// TwinCAT 3 PLC project TestRunner
// Title: TestRunner
// Company: Intecre Ltd
// ProjectVersion: 1.0.0.0
// Description: TcUnit test suites for the Intecre.Utilities library. Not a library; activate it on a runtime (the usermode runtime works) to run the tests.
// ProgramVersion: 3.1.4026.25
// libraries:
//   Tc2_Standard, * (Beckhoff Automation GmbH)
//   Tc2_System, * (Beckhoff Automation GmbH)
//   Tc2_Utilities, * (Beckhoff Automation GmbH)
//   TcUnit, * (www.tcunit.org)
//   Intecre.Utilities, * (Intecre Ltd)
// project tree:
//   / MAIN.TcPOU, PlcTask.TcTTO, SlowTask.TcTTO, ControllersInSlowTask.TcPOU
//   Tests/ CharIsNumber_Tests.TcPOU, TryStringToDint_Tests.TcPOU, TryStringToUdint_Tests.TcPOU, TryStringToWord_Tests.TcPOU, TryStringToLreal_Tests.TcPOU, F_Concat_Tests.TcPOU, F_ConcatLarge_Tests.TcPOU, F_Gate_Tests.TcPOU, FB_StringList_Tests.TcPOU, FB_UdintList_Tests.TcPOU, FB_PointerList_Tests.TcPOU, FB_LongStringList_Tests.TcPOU, FB_TargList_Tests.TcPOU, FB_Dictionary_Tests.TcPOU, F_DictionaryValuesCrc_Tests.TcPOU, FB_AlphaBetaFilter_Tests.TcPOU, FB_P_Control_Tests.TcPOU, FB_I_Controller_Tests.TcPOU, FB_PI_Controller_Tests.TcPOU, T_Task_Tests.TcPOU, T_NamedBase_Tests.TcPOU, Logger_Tests.TcPOU, FB_Assert_Tests.TcPOU, F_GetKL306xState_Tests.TcPOU, ProjectInformation_Tests.TcPOU, F_TargToString_Tests.TcPOU, F_StringToTarg_Tests.TcPOU, F_GetAmsNetId_Tests.TcPOU, T_Timer_Tests.TcPOU, T_GetHandle_Tests.TcPOU, T_InvokeRpcMethod_Tests.TcPOU, T_WritePersistentData_Tests.TcPOU
//   Mocks/ T_MockExternalLogger.TcPOU, T_RpcTarget.TcPOU, ST_RpcAddParams.TcDUT
// (motion and I/O tree: see PLC project intecreutilities)
// real-time tasks:
//   TASK PlcTask: cycle T#10ms, priority 20, ADS port 350
//   TASK SlowTask: cycle T#50000us, priority 25, ADS port 351

CONFIGURATION TestRunner
    RESOURCE PLC ON TwinCAT3
        TASK PlcTask(INTERVAL := T#10ms, PRIORITY := 20);
        TASK SlowTask(INTERVAL := T#50000us, PRIORITY := 25);
        PROGRAM MAIN WITH PlcTask : MAIN;
        PROGRAM ControllersInSlowTask WITH SlowTask : ControllersInSlowTask;
    END_RESOURCE
END_CONFIGURATION

// ---- Mocks/ST_RpcAddParams.TcDUT
// Input block of T_RpcTarget.Add as sent over ADS.
TYPE ST_RpcAddParams :
STRUCT
  a : DINT;
  b : DINT;
END_STRUCT
END_TYPE

// ---- MAIN.TcPOU
// Runs every TcUnit suite of the Intecre.Utilities library, one suite at a time.
PROGRAM MAIN
VAR
  suiteCharIsNumber        : CharIsNumber_Tests;
  suiteTryStringToDint     : TryStringToDint_Tests;
  suiteTryStringToUdint    : TryStringToUdint_Tests;
  suiteTryStringToWord     : TryStringToWord_Tests;
  suiteTryStringToLreal    : TryStringToLreal_Tests;
  suiteConcat              : F_Concat_Tests;
  suiteConcatLarge         : F_ConcatLarge_Tests;
  suiteGate                : F_Gate_Tests;
  suiteStringList          : FB_StringList_Tests;
  suiteUdintList           : FB_UdintList_Tests;
  suitePointerList         : FB_PointerList_Tests;
  suiteLongStringList      : FB_LongStringList_Tests;
  suiteTargList            : FB_TargList_Tests;
  suiteDictionary          : FB_Dictionary_Tests;
  suiteDictionaryValuesCrc : F_DictionaryValuesCrc_Tests;
  suiteAlphaBetaFilter     : FB_AlphaBetaFilter_Tests;
  suiteP_Control           : FB_P_Control_Tests;
  suiteI_Controller        : FB_I_Controller_Tests;
  suitePI_Controller       : FB_PI_Controller_Tests;
  suiteTask                : T_Task_Tests;
  suiteNamedBase           : T_NamedBase_Tests;
  suiteLogger              : Logger_Tests;
  suiteAssert              : FB_Assert_Tests;
  suiteGetKL306xState      : F_GetKL306xState_Tests;
  suiteProjectInformation  : ProjectInformation_Tests;
  suiteTargToString        : F_TargToString_Tests;
  suiteStringToTarg        : F_StringToTarg_Tests;
  suiteGetAmsNetId         : F_GetAmsNetId_Tests;
  suiteTimer               : T_Timer_Tests;
  suiteGetHandle           : T_GetHandle_Tests;
  suiteInvokeRpc           : T_InvokeRpcMethod_Tests;
  suiteWritePersistentData : T_WritePersistentData_Tests;
END_VAR

TcUnit.RUN_IN_SEQUENCE();

END_PROGRAM

// ---- Tests/CharIsNumber_Tests.TcPOU
FUNCTION_BLOCK CharIsNumber_Tests EXTENDS TcUnit.FB_TestSuite

Test_DigitsAreNumbers();
Test_NonDigitsAreNotNumbers();
Test_MinusAcceptedOnlyByOrMinus();
Test_PeriodAcceptedOnlyByOrPeriod();

METHOD PRIVATE Test_DigitsAreNumbers
VAR
  ch : BYTE;
  allDigits : BOOL := TRUE;
END_VAR
TcUnit.TEST(__POUNAME());

// arrange / act
FOR ch := 48 TO 57 DO
  allDigits := allDigits AND CharIsNumber(ch);
END_FOR

// assert
AssertTrue(Condition := allDigits, Message := 'ASCII 0-9 are numbers');

TEST_FINISHED_NAMED(__POUNAME());
END_METHOD

METHOD PRIVATE Test_NonDigitsAreNotNumbers
TcUnit.TEST(__POUNAME());

// act / assert
AssertFalse(Condition := CharIsNumber(47), Message := 'slash (47) is not a number');
AssertFalse(Condition := CharIsNumber(58), Message := 'colon (58) is not a number');
AssertFalse(Condition := CharIsNumber(65), Message := 'A is not a number');
AssertFalse(Condition := CharIsNumber(32), Message := 'space is not a number');
AssertFalse(Condition := CharIsNumber(45), Message := 'minus is not a number');
AssertFalse(Condition := CharIsNumber(46), Message := 'period is not a number');

TEST_FINISHED_NAMED(__POUNAME());
END_METHOD

METHOD PRIVATE Test_MinusAcceptedOnlyByOrMinus
TcUnit.TEST(__POUNAME());

// act / assert
AssertTrue(Condition := CharIsNumberOrMinus(45), Message := 'minus accepted');
AssertTrue(Condition := CharIsNumberOrMinus(53), Message := 'digit 5 accepted');
AssertFalse(Condition := CharIsNumberOrMinus(46), Message := 'period rejected');
AssertFalse(Condition := CharIsNumberOrMinus(65), Message := 'letter rejected');

TEST_FINISHED_NAMED(__POUNAME());
END_METHOD

METHOD PRIVATE Test_PeriodAcceptedOnlyByOrPeriod
TcUnit.TEST(__POUNAME());

// act / assert
AssertTrue(Condition := CharIsNumberOrPeriod(46), Message := 'period accepted');
AssertTrue(Condition := CharIsNumberOrPeriod(48), Message := 'digit 0 accepted');
AssertFalse(Condition := CharIsNumberOrPeriod(45), Message := 'minus rejected');
AssertFalse(Condition := CharIsNumberOrPeriod(65), Message := 'letter rejected');

TEST_FINISHED_NAMED(__POUNAME());
END_METHOD

END_FUNCTION_BLOCK

// ---- Tests/TryStringToDint_Tests.TcPOU
FUNCTION_BLOCK TryStringToDint_Tests EXTENDS TcUnit.FB_TestSuite

Test_ParsesPositive();
Test_ParsesNegative();
Test_ParsesMaxValue();
Test_RejectsLetters();
Test_RejectsEmptyString();
Test_RejectsMinusInsideNumber();
Test_RejectsPlusSign();

METHOD PRIVATE Test_ParsesPositive
VAR
  value : DINT;
  ok : BOOL;
END_VAR
TcUnit.TEST(__POUNAME());

// act
ok := TryStringToDint('123', value);

// assert
AssertTrue(Condition := ok, Message := '123 parses');
AssertEquals_DINT(Expected := 123, Actual := value, Message := 'parsed value');

TEST_FINISHED_NAMED(__POUNAME());
END_METHOD

METHOD PRIVATE Test_ParsesNegative
VAR
  value : DINT;
  ok : BOOL;
END_VAR
TcUnit.TEST(__POUNAME());

// act
ok := TryStringToDint('-45', value);

// assert
AssertTrue(Condition := ok, Message := '-45 parses');
AssertEquals_DINT(Expected := -45, Actual := value, Message := 'parsed value');

TEST_FINISHED_NAMED(__POUNAME());
END_METHOD

METHOD PRIVATE Test_ParsesMaxValue
VAR
  value : DINT;
  ok : BOOL;
END_VAR
TcUnit.TEST(__POUNAME());

// act
ok := TryStringToDint('2147483647', value);

// assert
AssertTrue(Condition := ok, Message := 'DINT max parses');
AssertEquals_DINT(Expected := 2147483647, Actual := value, Message := 'parsed value');

TEST_FINISHED_NAMED(__POUNAME());
END_METHOD

METHOD PRIVATE Test_RejectsLetters
VAR
  value : DINT;
  ok : BOOL;
END_VAR
TcUnit.TEST(__POUNAME());

// arrange
value := 99;

// act
ok := TryStringToDint('12a', value);

// assert
AssertFalse(Condition := ok, Message := 'letters rejected');
AssertEquals_DINT(Expected := 0, Actual := value, Message := 'value cleared on failure');

TEST_FINISHED_NAMED(__POUNAME());
END_METHOD

METHOD PRIVATE Test_RejectsEmptyString
VAR
  value : DINT;
  ok : BOOL;
END_VAR
TcUnit.TEST(__POUNAME());

// arrange
value := 99;

// act
ok := TryStringToDint('', value);

// assert
AssertFalse(Condition := ok, Message := 'empty string rejected');
AssertEquals_DINT(Expected := 0, Actual := value, Message := 'value cleared on failure');

TEST_FINISHED_NAMED(__POUNAME());
END_METHOD

METHOD PRIVATE Test_RejectsMinusInsideNumber
VAR
  value : DINT;
  ok : BOOL;
END_VAR
TcUnit.TEST(__POUNAME());

// act
ok := TryStringToDint('1-2', value);

// assert
AssertFalse(Condition := ok, Message := 'minus only allowed as first character');

TEST_FINISHED_NAMED(__POUNAME());
END_METHOD

METHOD PRIVATE Test_RejectsPlusSign
VAR
  value : DINT;
  ok : BOOL;
END_VAR
TcUnit.TEST(__POUNAME());

// act
ok := TryStringToDint('+1', value);

// assert
AssertFalse(Condition := ok, Message := 'explicit plus sign is not accepted');

TEST_FINISHED_NAMED(__POUNAME());
END_METHOD

END_FUNCTION_BLOCK

// ---- Tests/TryStringToUdint_Tests.TcPOU
FUNCTION_BLOCK TryStringToUdint_Tests EXTENDS TcUnit.FB_TestSuite

Test_ParsesZero();
Test_ParsesMaxValue();
Test_RejectsNegative();
Test_RejectsEmptyString();
Test_RejectsTrailingSpace();

METHOD PRIVATE Test_ParsesZero
VAR
  value : UDINT;
  ok : BOOL;
END_VAR
TcUnit.TEST(__POUNAME());

// act
ok := TryStringToUdint('0', value);

// assert
AssertTrue(Condition := ok, Message := '0 parses');
AssertEquals_UDINT(Expected := 0, Actual := value, Message := 'parsed value');

TEST_FINISHED_NAMED(__POUNAME());
END_METHOD

METHOD PRIVATE Test_ParsesMaxValue
VAR
  value : UDINT;
  ok : BOOL;
END_VAR
TcUnit.TEST(__POUNAME());

// act
ok := TryStringToUdint('4294967295', value);

// assert
AssertTrue(Condition := ok, Message := 'UDINT max parses');
AssertEquals_UDINT(Expected := 4294967295, Actual := value, Message := 'parsed value');

TEST_FINISHED_NAMED(__POUNAME());
END_METHOD

METHOD PRIVATE Test_RejectsNegative
VAR
  value : UDINT;
  ok : BOOL;
END_VAR
TcUnit.TEST(__POUNAME());

// arrange
value := 99;

// act
ok := TryStringToUdint('-1', value);

// assert
AssertFalse(Condition := ok, Message := 'negative rejected');
AssertEquals_UDINT(Expected := 0, Actual := value, Message := 'value cleared on failure');

TEST_FINISHED_NAMED(__POUNAME());
END_METHOD

METHOD PRIVATE Test_RejectsEmptyString
VAR
  value : UDINT;
  ok : BOOL;
END_VAR
TcUnit.TEST(__POUNAME());

// arrange
value := 99;

// act
ok := TryStringToUdint('', value);

// assert
AssertFalse(Condition := ok, Message := 'empty string rejected');
AssertEquals_UDINT(Expected := 0, Actual := value, Message := 'value cleared on failure');

TEST_FINISHED_NAMED(__POUNAME());
END_METHOD

METHOD PRIVATE Test_RejectsTrailingSpace
VAR
  value : UDINT;
  ok : BOOL;
END_VAR
TcUnit.TEST(__POUNAME());

// act
ok := TryStringToUdint('12 ', value);

// assert
AssertFalse(Condition := ok, Message := 'trailing space rejected');

TEST_FINISHED_NAMED(__POUNAME());
END_METHOD

END_FUNCTION_BLOCK

// ---- Tests/TryStringToWord_Tests.TcPOU
FUNCTION_BLOCK TryStringToWord_Tests EXTENDS TcUnit.FB_TestSuite

Test_ParsesValue();
Test_ParsesMaxValue();
Test_RejectsOverflow();
Test_RejectsLetters();

METHOD PRIVATE Test_ParsesValue
VAR
  value : WORD;
  ok : BOOL;
END_VAR
TcUnit.TEST(__POUNAME());

// act
ok := TryStringToWord('7', value);

// assert
AssertTrue(Condition := ok, Message := '7 parses');
AssertEquals_WORD(Expected := 7, Actual := value, Message := 'parsed value');

TEST_FINISHED_NAMED(__POUNAME());
END_METHOD

METHOD PRIVATE Test_ParsesMaxValue
VAR
  value : WORD;
  ok : BOOL;
END_VAR
TcUnit.TEST(__POUNAME());

// act
ok := TryStringToWord('65535', value);

// assert
AssertTrue(Condition := ok, Message := 'WORD max parses');
AssertEquals_WORD(Expected := 65535, Actual := value, Message := 'parsed value');

TEST_FINISHED_NAMED(__POUNAME());
END_METHOD

METHOD PRIVATE Test_RejectsOverflow
VAR
  value : WORD;
  ok : BOOL;
END_VAR
TcUnit.TEST(__POUNAME());

// arrange
value := 99;

// act
ok := TryStringToWord('65536', value);

// assert
AssertFalse(Condition := ok, Message := '65536 does not fit a WORD');
AssertEquals_WORD(Expected := 0, Actual := value, Message := 'value cleared on failure');

TEST_FINISHED_NAMED(__POUNAME());
END_METHOD

METHOD PRIVATE Test_RejectsLetters
VAR
  value : WORD;
  ok : BOOL;
END_VAR
TcUnit.TEST(__POUNAME());

// act
ok := TryStringToWord('abc', value);

// assert
AssertFalse(Condition := ok, Message := 'letters rejected');

TEST_FINISHED_NAMED(__POUNAME());
END_METHOD

END_FUNCTION_BLOCK

// ---- Tests/TryStringToLreal_Tests.TcPOU
FUNCTION_BLOCK TryStringToLreal_Tests EXTENDS TcUnit.FB_TestSuite

Test_ParsesDecimal();
Test_ParsesNegativeDecimal();
Test_ParsesInteger();
Test_ParsesNegativeFraction();
Test_ParsesSmallFraction();
Test_RejectsLetters();
Test_RejectsExponent();
Test_RejectsEmptyString();

METHOD PRIVATE Test_ParsesDecimal
VAR
  value : LREAL;
  ok : BOOL;
END_VAR
TcUnit.TEST(__POUNAME());

// act
ok := TryStringToLreal('3.25', value);

// assert
AssertTrue(Condition := ok, Message := '3.25 parses');
AssertEquals_LREAL(Expected := 3.25, Actual := value, Delta := 1.0E-9, Message := 'parsed value');

TEST_FINISHED_NAMED(__POUNAME());
END_METHOD

METHOD PRIVATE Test_ParsesNegativeDecimal
VAR
  value : LREAL;
  ok : BOOL;
END_VAR
TcUnit.TEST(__POUNAME());

// act
ok := TryStringToLreal('-1.5', value);

// assert
AssertTrue(Condition := ok, Message := '-1.5 parses');
AssertEquals_LREAL(Expected := -1.5, Actual := value, Delta := 1.0E-9, Message := 'sign applies to the whole number');

TEST_FINISHED_NAMED(__POUNAME());
END_METHOD

METHOD PRIVATE Test_ParsesInteger
VAR
  value : LREAL;
  ok : BOOL;
END_VAR
TcUnit.TEST(__POUNAME());

// act
ok := TryStringToLreal('42', value);

// assert
AssertTrue(Condition := ok, Message := '42 parses');
AssertEquals_LREAL(Expected := 42.0, Actual := value, Delta := 1.0E-9, Message := 'integer text parses as LREAL');

TEST_FINISHED_NAMED(__POUNAME());
END_METHOD

METHOD PRIVATE Test_ParsesNegativeFraction
VAR
  value : LREAL;
  ok : BOOL;
END_VAR
TcUnit.TEST(__POUNAME());

// act
ok := TryStringToLreal('-0.5', value);

// assert
AssertTrue(Condition := ok, Message := '-0.5 parses');
AssertEquals_LREAL(Expected := -0.5, Actual := value, Delta := 1.0E-9, Message := 'sign kept when the integer part is zero');

TEST_FINISHED_NAMED(__POUNAME());
END_METHOD

METHOD PRIVATE Test_ParsesSmallFraction
VAR
  value : LREAL;
  ok : BOOL;
END_VAR
TcUnit.TEST(__POUNAME());

// act
ok := TryStringToLreal('0.001', value);

// assert
AssertTrue(Condition := ok, Message := '0.001 parses');
AssertEquals_LREAL(Expected := 0.001, Actual := value, Delta := 1.0E-9, Message := 'leading zeros in the fraction are kept');

TEST_FINISHED_NAMED(__POUNAME());
END_METHOD

METHOD PRIVATE Test_RejectsLetters
VAR
  value : LREAL;
  ok : BOOL;
END_VAR
TcUnit.TEST(__POUNAME());

// arrange
value := 9.9;

// act
ok := TryStringToLreal('abc', value);

// assert
AssertFalse(Condition := ok, Message := 'letters rejected');
AssertEquals_LREAL(Expected := 0.0, Actual := value, Delta := 1.0E-9, Message := 'value cleared on failure');

TEST_FINISHED_NAMED(__POUNAME());
END_METHOD

METHOD PRIVATE Test_RejectsExponent
VAR
  value : LREAL;
  ok : BOOL;
END_VAR
TcUnit.TEST(__POUNAME());

// act
ok := TryStringToLreal('1e5', value);

// assert
AssertFalse(Condition := ok, Message := 'exponent notation rejected');

TEST_FINISHED_NAMED(__POUNAME());
END_METHOD

METHOD PRIVATE Test_RejectsEmptyString
VAR
  value : LREAL;
  ok : BOOL;
END_VAR
TcUnit.TEST(__POUNAME());

// arrange
value := 9.9;

// act
ok := TryStringToLreal('', value);

// assert
AssertFalse(Condition := ok, Message := 'empty string rejected');
AssertEquals_LREAL(Expected := 0.0, Actual := value, Delta := 1.0E-9, Message := 'value cleared on failure');

TEST_FINISHED_NAMED(__POUNAME());
END_METHOD

END_FUNCTION_BLOCK

// ---- Tests/F_Concat_Tests.TcPOU
FUNCTION_BLOCK F_Concat_Tests EXTENDS TcUnit.FB_TestSuite

Test_Concat3();
Test_Concat4();
Test_Concat5();
Test_Concat6();
Test_Concat7();
Test_EmptyPartsAreSkipped();
Test_ResultLimitedToMaxString();

METHOD PRIVATE Test_Concat3
TcUnit.TEST(__POUNAME());

AssertEquals_STRING(Expected := 'abc', Actual := F_Concat3('a', 'b', 'c'), Message := 'three parts joined');

TEST_FINISHED_NAMED(__POUNAME());
END_METHOD

METHOD PRIVATE Test_Concat4
TcUnit.TEST(__POUNAME());

AssertEquals_STRING(Expected := 'abcd', Actual := F_Concat4('a', 'b', 'c', 'd'), Message := 'four parts joined');

TEST_FINISHED_NAMED(__POUNAME());
END_METHOD

METHOD PRIVATE Test_Concat5
TcUnit.TEST(__POUNAME());

AssertEquals_STRING(Expected := 'abcde', Actual := F_Concat5('a', 'b', 'c', 'd', 'e'), Message := 'five parts joined');

TEST_FINISHED_NAMED(__POUNAME());
END_METHOD

METHOD PRIVATE Test_Concat6
TcUnit.TEST(__POUNAME());

AssertEquals_STRING(Expected := 'abcdef', Actual := F_Concat6('a', 'b', 'c', 'd', 'e', 'f'), Message := 'six parts joined');

TEST_FINISHED_NAMED(__POUNAME());
END_METHOD

METHOD PRIVATE Test_Concat7
TcUnit.TEST(__POUNAME());

AssertEquals_STRING(Expected := 'abcdefg', Actual := F_Concat7('a', 'b', 'c', 'd', 'e', 'f', 'g'), Message := 'seven parts joined');

TEST_FINISHED_NAMED(__POUNAME());
END_METHOD

METHOD PRIVATE Test_EmptyPartsAreSkipped
TcUnit.TEST(__POUNAME());

AssertEquals_STRING(Expected := 'x', Actual := F_Concat3('', 'x', ''), Message := 'empty parts contribute nothing');

TEST_FINISHED_NAMED(__POUNAME());
END_METHOD

METHOD PRIVATE Test_ResultLimitedToMaxString
VAR
  part : STRING;
  i : INT;
  result : T_MaxString;
END_VAR
TcUnit.TEST(__POUNAME());

// arrange
FOR i := 1 TO 80 DO
  part := CONCAT(part, 'x');
END_FOR

// act
result := F_Concat4(part, part, part, part);

// assert
AssertEquals_INT(Expected := 255, Actual := LEN(result), Message := '4 x 80 characters truncate to T_MaxString');

TEST_FINISHED_NAMED(__POUNAME());
END_METHOD

END_FUNCTION_BLOCK

// ---- Tests/F_ConcatLarge_Tests.TcPOU
FUNCTION_BLOCK F_ConcatLarge_Tests EXTENDS TcUnit.FB_TestSuite
VAR
  one, two, three, four, five, six, seven : LongString;
  result : LongString;
END_VAR

Test_ConcatsTwoStrings();
Test_TruncatesFirstStringToFitMaxLength();
Test_Concat3Large();
Test_Concat4Large();
Test_Concat5Large();
Test_Concat6Large();
Test_Concat7Large();
Test_ClearLargeEmptiesString();

// Test helper: a LongString of count copies of the byte ch.
METHOD PRIVATE Fill : LongString
VAR_INPUT
  count : INT;
  ch : BYTE;
END_VAR
VAR
  i : INT;
  text : LongString;
END_VAR
FOR i := 0 TO count - 1 DO
  text[i] := ch;
END_FOR
text[count] := 0;
Fill := text;
END_METHOD

METHOD PRIVATE Test_ClearLargeEmptiesString
TcUnit.TEST(__POUNAME());

// arrange
one := 'abc';

// act
F_ClearLarge(one);

// assert
AssertEquals_INT(Expected := 0, Actual := LEN(one), Message := 'cleared string is empty');
AssertEquals_BYTE(Expected := 0, Actual := one[1], Message := 'bytes behind the terminator are zeroed too');

TEST_FINISHED_NAMED(__POUNAME());
END_METHOD

METHOD PRIVATE Test_Concat3Large
TcUnit.TEST(__POUNAME());

one := 'a'; two := 'b'; three := 'c';
result := F_Concat3_Large(one, two, three);
AssertTrue(Condition := result = 'abc', Message := 'three long strings joined');

TEST_FINISHED_NAMED(__POUNAME());
END_METHOD

METHOD PRIVATE Test_Concat4Large
TcUnit.TEST(__POUNAME());

one := 'a'; two := 'b'; three := 'c'; four := 'd';
result := F_Concat4_Large(one, two, three, four);
AssertTrue(Condition := result = 'abcd', Message := 'four long strings joined');

TEST_FINISHED_NAMED(__POUNAME());
END_METHOD

METHOD PRIVATE Test_Concat5Large
TcUnit.TEST(__POUNAME());

one := 'a'; two := 'b'; three := 'c'; four := 'd'; five := 'e';
result := F_Concat5_Large(one, two, three, four, five);
AssertTrue(Condition := result = 'abcde', Message := 'five long strings joined');

TEST_FINISHED_NAMED(__POUNAME());
END_METHOD

METHOD PRIVATE Test_Concat6Large
TcUnit.TEST(__POUNAME());

one := 'a'; two := 'b'; three := 'c'; four := 'd'; five := 'e'; six := 'f';
result := F_Concat6_Large(one, two, three, four, five, six);
AssertTrue(Condition := result = 'abcdef', Message := 'six long strings joined');

TEST_FINISHED_NAMED(__POUNAME());
END_METHOD

METHOD PRIVATE Test_Concat7Large
TcUnit.TEST(__POUNAME());

one := 'a'; two := 'b'; three := 'c'; four := 'd'; five := 'e'; six := 'f'; seven := 'g';
result := F_Concat7_Large(one, two, three, four, five, six, seven);
AssertTrue(Condition := result = 'abcdefg', Message := 'seven long strings joined');

TEST_FINISHED_NAMED(__POUNAME());
END_METHOD

METHOD PRIVATE Test_ConcatsTwoStrings
TcUnit.TEST(__POUNAME());

// arrange
one := 'abc';
two := 'def';

// act
result := F_ConcatLarge(one, two);

// assert
AssertTrue(Condition := result = 'abcdef', Message := 'two long strings joined');
AssertEquals_INT(Expected := 6, Actual := LEN(result), Message := 'length of the join');

TEST_FINISHED_NAMED(__POUNAME());
END_METHOD

METHOD PRIVATE Test_TruncatesFirstStringToFitMaxLength
TcUnit.TEST(__POUNAME());

// arrange: 150 + 150 characters exceed the 299 usable characters of a LongString
one := Fill(150, 97); // 'a'
two := Fill(150, 98); // 'b'

// act
result := F_ConcatLarge(one, two);

// assert (LEN stops at 255 characters, LEN2 measures the whole string)
AssertEquals_UDINT(Expected := 299, Actual := LEN2(ADR(result)), Message := 'result fills the LongString');
AssertEquals_BYTE(Expected := 97, Actual := result[148], Message := 'first string keeps 149 characters');
AssertEquals_BYTE(Expected := 98, Actual := result[149], Message := 'second string starts where the first was cut');
AssertEquals_BYTE(Expected := 98, Actual := result[298], Message := 'second string kept whole');
AssertEquals_BYTE(Expected := 0, Actual := result[299], Message := 'terminator in the last position');

// arrange: a second string longer than 255 characters must be measured in full
one := Fill(10, 97);
two := Fill(280, 98);

// act
result := F_ConcatLarge(one, two);

// assert
AssertEquals_UDINT(Expected := 290, Actual := LEN2(ADR(result)), Message := 'inputs over 255 characters are measured in full');
AssertEquals_BYTE(Expected := 97, Actual := result[9], Message := 'first string copied whole');
AssertEquals_BYTE(Expected := 98, Actual := result[289], Message := 'last character of the second string kept');
AssertEquals_BYTE(Expected := 0, Actual := result[290], Message := 'terminator after the join');

TEST_FINISHED_NAMED(__POUNAME());
END_METHOD

END_FUNCTION_BLOCK

// ---- Tests/F_Gate_Tests.TcPOU
FUNCTION_BLOCK F_Gate_Tests EXTENDS TcUnit.FB_TestSuite

Test_ReturnsTrueAndResetsFlag();
Test_ReturnsFalseWhenFlagClear();

METHOD PRIVATE Test_ReturnsTrueAndResetsFlag
VAR
  flag : BOOL;
  result : BOOL;
END_VAR
TcUnit.TEST(__POUNAME());

// arrange
flag := TRUE;

// act
result := F_Gate(flag);

// assert
AssertTrue(Condition := result, Message := 'returns the flag as it was');
AssertFalse(Condition := flag, Message := 'flag reset by the call');

TEST_FINISHED_NAMED(__POUNAME());
END_METHOD

METHOD PRIVATE Test_ReturnsFalseWhenFlagClear
VAR
  flag : BOOL;
  result : BOOL;
END_VAR
TcUnit.TEST(__POUNAME());

// arrange
flag := FALSE;

// act
result := F_Gate(flag);

// assert
AssertFalse(Condition := result, Message := 'clear flag reads FALSE');
AssertFalse(Condition := flag, Message := 'flag stays clear');

TEST_FINISHED_NAMED(__POUNAME());
END_METHOD

END_FUNCTION_BLOCK

// ---- Tests/FB_StringList_Tests.TcPOU
FUNCTION_BLOCK FB_StringList_Tests EXTENDS TcUnit.FB_TestSuite
VAR
  list : FB_StringList;
  copy : ARRAY[0..GVL_List.LIST_SIZE - 1] OF T_MaxString;
END_VAR

Test_AddItemIncrementsCount();
Test_ContainsFindsAddedItem();
Test_FindIndexReturnsPosition();
Test_GetIndexReturnsItem();
Test_TryGetIndexLeavesItemOnFailure();
Test_RemoveIndexShiftsItems();
Test_RemoveIndexRejectsOutOfRange();
Test_GetAndRemoveIndex();
Test_ClearEmptiesList();
Test_RejectsAddWhenFull();
Test_ContainsPartialMatchesSubstring();
Test_CopyListAndClearCopiesThenEmpties();

METHOD PRIVATE Test_AddItemIncrementsCount
VAR
  ok : BOOL;
END_VAR
TcUnit.TEST(__POUNAME());

// arrange
list.Clear();

// act
ok := list.AddItem('one');

// assert
AssertTrue(Condition := ok, Message := 'add succeeds');
AssertEquals_UDINT(Expected := 1, Actual := list.Count, Message := 'count after one add');

TEST_FINISHED_NAMED(__POUNAME());
END_METHOD

METHOD PRIVATE Test_ContainsFindsAddedItem
TcUnit.TEST(__POUNAME());

// arrange
list.Clear();
list.AddItem('one');
list.AddItem('two');

// assert
AssertTrue(Condition := list.Contains('two'), Message := 'added item found');
AssertFalse(Condition := list.Contains('three'), Message := 'missing item not found');

TEST_FINISHED_NAMED(__POUNAME());
END_METHOD

METHOD PRIVATE Test_FindIndexReturnsPosition
TcUnit.TEST(__POUNAME());

// arrange
list.Clear();
list.AddItem('a');
list.AddItem('b');
list.AddItem('c');

// assert
AssertEquals_INT(Expected := 2, Actual := list.FindIndex('c'), Message := 'index of the third item');
AssertEquals_INT(Expected := -1, Actual := list.FindIndex('zzz'), Message := 'missing item gives -1');

TEST_FINISHED_NAMED(__POUNAME());
END_METHOD

METHOD PRIVATE Test_GetIndexReturnsItem
TcUnit.TEST(__POUNAME());

// arrange
list.Clear();
list.AddItem('a');
list.AddItem('b');

// assert
AssertEquals_STRING(Expected := 'b', Actual := list.GetIndex(1), Message := 'item at index 1');
AssertEquals_STRING(Expected := '', Actual := list.GetIndex(5), Message := 'out of range gives empty');

TEST_FINISHED_NAMED(__POUNAME());
END_METHOD

METHOD PRIVATE Test_TryGetIndexLeavesItemOnFailure
VAR
  ok : BOOL;
  item : T_MaxString;
END_VAR
TcUnit.TEST(__POUNAME());

// arrange
list.Clear();
list.AddItem('a');
item := 'unchanged';

// act
ok := list.TryGetIndex(5, item);

// assert
AssertFalse(Condition := ok, Message := 'out of range fails');
AssertEquals_STRING(Expected := 'unchanged', Actual := item, Message := 'item untouched');

TEST_FINISHED_NAMED(__POUNAME());
END_METHOD

METHOD PRIVATE Test_RemoveIndexShiftsItems
VAR
  ok : BOOL;
END_VAR
TcUnit.TEST(__POUNAME());

// arrange
list.Clear();
list.AddItem('a');
list.AddItem('b');
list.AddItem('c');

// act
ok := list.RemoveIndex(1);

// assert
AssertTrue(Condition := ok, Message := 'remove succeeds');
AssertEquals_UDINT(Expected := 2, Actual := list.Count, Message := 'count after remove');
AssertEquals_STRING(Expected := 'a', Actual := list.GetIndex(0), Message := 'first item kept');
AssertEquals_STRING(Expected := 'c', Actual := list.GetIndex(1), Message := 'last item shifted down');
AssertEquals_STRING(Expected := '', Actual := list.GetIndex(2), Message := 'old slot cleared');

TEST_FINISHED_NAMED(__POUNAME());
END_METHOD

METHOD PRIVATE Test_RemoveIndexRejectsOutOfRange
VAR
  ok : BOOL;
END_VAR
TcUnit.TEST(__POUNAME());

// arrange
list.Clear();
list.AddItem('a');

// act
ok := list.RemoveIndex(1);

// assert
AssertFalse(Condition := ok, Message := 'out of range rejected');
AssertEquals_UDINT(Expected := 1, Actual := list.Count, Message := 'count unchanged');

TEST_FINISHED_NAMED(__POUNAME());
END_METHOD

METHOD PRIVATE Test_GetAndRemoveIndex
VAR
  item : T_MaxString;
END_VAR
TcUnit.TEST(__POUNAME());

// arrange
list.Clear();
list.AddItem('a');
list.AddItem('b');

// act
item := list.GetAndRemoveIndex(0);

// assert
AssertEquals_STRING(Expected := 'a', Actual := item, Message := 'removed item returned');
AssertEquals_UDINT(Expected := 1, Actual := list.Count, Message := 'count after remove');
AssertEquals_STRING(Expected := 'b', Actual := list.GetIndex(0), Message := 'remaining item shifted down');

TEST_FINISHED_NAMED(__POUNAME());
END_METHOD

METHOD PRIVATE Test_ClearEmptiesList
TcUnit.TEST(__POUNAME());

// arrange
list.Clear();
list.AddItem('a');
list.AddItem('b');

// act
list.Clear();

// assert
AssertEquals_UDINT(Expected := 0, Actual := list.Count, Message := 'count after clear');
AssertFalse(Condition := list.Contains('a'), Message := 'items gone after clear');

TEST_FINISHED_NAMED(__POUNAME());
END_METHOD

METHOD PRIVATE Test_RejectsAddWhenFull
VAR
  i : UINT;
  ok : BOOL;
END_VAR
TcUnit.TEST(__POUNAME());

// arrange
list.Clear();
FOR i := 1 TO GVL_List.LIST_SIZE DO
  list.AddItem(CONCAT('item', TO_STRING(i)));
END_FOR

// act
ok := list.AddItem('overflow');

// assert
AssertEquals_UDINT(Expected := TO_UDINT(GVL_List.LIST_SIZE), Actual := list.Count, Message := 'list holds LIST_SIZE items');
AssertFalse(Condition := ok, Message := 'add rejected when full');

TEST_FINISHED_NAMED(__POUNAME());
END_METHOD

METHOD PRIVATE Test_ContainsPartialMatchesSubstring
TcUnit.TEST(__POUNAME());

// arrange
list.Clear();
list.AddItem('hello world');

// assert
AssertTrue(Condition := list.ContainsPartial('lo wo'), Message := 'substring found');
AssertFalse(Condition := list.ContainsPartial('xyz'), Message := 'missing substring not found');
AssertEquals_INT(Expected := 0, Actual := list.FindIndexPartialKey('world'), Message := 'index of the partial match');

TEST_FINISHED_NAMED(__POUNAME());
END_METHOD

METHOD PRIVATE Test_CopyListAndClearCopiesThenEmpties
TcUnit.TEST(__POUNAME());

// arrange
list.Clear();
list.AddItem('a');
list.AddItem('b');

// act
list.CopyListAndClear(copy);

// assert
AssertEquals_STRING(Expected := 'a', Actual := copy[0], Message := 'first item copied');
AssertEquals_STRING(Expected := 'b', Actual := copy[1], Message := 'second item copied');
AssertEquals_UDINT(Expected := 0, Actual := list.Count, Message := 'list emptied');

TEST_FINISHED_NAMED(__POUNAME());
END_METHOD

END_FUNCTION_BLOCK

// ---- Tests/FB_UdintList_Tests.TcPOU
FUNCTION_BLOCK FB_UdintList_Tests EXTENDS TcUnit.FB_TestSuite
VAR
  list : FB_UdintList;
END_VAR

Test_AddItemIncrementsCount();
Test_ContainsFindsAddedItem();
Test_FindIndexReturnsPosition();
Test_GetIndexReturnsItem();
Test_TryGetIndexClearsItemOnFailure();
Test_RemoveIndexShiftsItems();
Test_ClearEmptiesList();
Test_RejectsAddWhenFull();

METHOD PRIVATE Test_AddItemIncrementsCount
VAR
  ok : BOOL;
END_VAR
TcUnit.TEST(__POUNAME());

list.Clear();
ok := list.AddItem(10);
AssertTrue(Condition := ok, Message := 'add succeeds');
AssertEquals_UDINT(Expected := 1, Actual := list.Count, Message := 'count after one add');

TEST_FINISHED_NAMED(__POUNAME());
END_METHOD

METHOD PRIVATE Test_ContainsFindsAddedItem
TcUnit.TEST(__POUNAME());

list.Clear();
list.AddItem(10);
list.AddItem(20);
AssertTrue(Condition := list.Contains(20), Message := 'added item found');
AssertFalse(Condition := list.Contains(30), Message := 'missing item not found');

TEST_FINISHED_NAMED(__POUNAME());
END_METHOD

METHOD PRIVATE Test_FindIndexReturnsPosition
TcUnit.TEST(__POUNAME());

list.Clear();
list.AddItem(10);
list.AddItem(20);
list.AddItem(30);
AssertEquals_INT(Expected := 2, Actual := list.FindIndex(30), Message := 'index of the third item');
AssertEquals_INT(Expected := -1, Actual := list.FindIndex(99), Message := 'missing item gives -1');

TEST_FINISHED_NAMED(__POUNAME());
END_METHOD

METHOD PRIVATE Test_GetIndexReturnsItem
TcUnit.TEST(__POUNAME());

list.Clear();
list.AddItem(10);
list.AddItem(20);
AssertEquals_UDINT(Expected := 20, Actual := list.GetIndex(1), Message := 'item at index 1');
AssertEquals_UDINT(Expected := 0, Actual := list.GetIndex(9), Message := 'out of range gives 0');

TEST_FINISHED_NAMED(__POUNAME());
END_METHOD

METHOD PRIVATE Test_TryGetIndexClearsItemOnFailure
VAR
  ok : BOOL;
  item : UDINT;
END_VAR
TcUnit.TEST(__POUNAME());

list.Clear();
list.AddItem(10);
item := 5;
ok := list.TryGetIndex(9, item);
AssertFalse(Condition := ok, Message := 'out of range fails');
AssertEquals_UDINT(Expected := 0, Actual := item, Message := 'item cleared to 0');

TEST_FINISHED_NAMED(__POUNAME());
END_METHOD

METHOD PRIVATE Test_RemoveIndexShiftsItems
VAR
  ok : BOOL;
END_VAR
TcUnit.TEST(__POUNAME());

list.Clear();
list.AddItem(10);
list.AddItem(20);
list.AddItem(30);
ok := list.RemoveIndex(1);
AssertTrue(Condition := ok, Message := 'remove succeeds');
AssertEquals_UDINT(Expected := 2, Actual := list.Count, Message := 'count after remove');
AssertEquals_UDINT(Expected := 10, Actual := list.GetIndex(0), Message := 'first item kept');
AssertEquals_UDINT(Expected := 30, Actual := list.GetIndex(1), Message := 'last item shifted down');
AssertFalse(Condition := list.RemoveIndex(7), Message := 'out of range rejected');

TEST_FINISHED_NAMED(__POUNAME());
END_METHOD

METHOD PRIVATE Test_ClearEmptiesList
TcUnit.TEST(__POUNAME());

list.Clear();
list.AddItem(10);
list.Clear();
AssertEquals_UDINT(Expected := 0, Actual := list.Count, Message := 'count after clear');
AssertFalse(Condition := list.Contains(10), Message := 'items gone after clear');

TEST_FINISHED_NAMED(__POUNAME());
END_METHOD

METHOD PRIVATE Test_RejectsAddWhenFull
VAR
  i : UINT;
  ok : BOOL;
END_VAR
TcUnit.TEST(__POUNAME());

list.Clear();
FOR i := 1 TO GVL_List.LIST_SIZE DO
  list.AddItem(i);
END_FOR
ok := list.AddItem(9999);
AssertEquals_UDINT(Expected := TO_UDINT(GVL_List.LIST_SIZE), Actual := list.Count, Message := 'list holds LIST_SIZE items');
AssertFalse(Condition := ok, Message := 'add rejected when full');

TEST_FINISHED_NAMED(__POUNAME());
END_METHOD

END_FUNCTION_BLOCK

// ---- Tests/FB_PointerList_Tests.TcPOU
FUNCTION_BLOCK FB_PointerList_Tests EXTENDS TcUnit.FB_TestSuite
VAR
  list : FB_PointerList;
  a, b, c : INT;
END_VAR

Test_AddAndContains();
Test_FindIndexReturnsPosition();
Test_GetIndexReturnsPointer();
Test_RemoveIndexShiftsItems();
Test_ClearEmptiesList();

METHOD PRIVATE Test_AddAndContains
TcUnit.TEST(__POUNAME());

list.Clear();
list.AddItem(ADR(a));
list.AddItem(ADR(b));
AssertEquals_UDINT(Expected := 2, Actual := list.Count, Message := 'count after two adds');
AssertTrue(Condition := list.Contains(ADR(b)), Message := 'added pointer found');
AssertFalse(Condition := list.Contains(ADR(c)), Message := 'missing pointer not found');

TEST_FINISHED_NAMED(__POUNAME());
END_METHOD

METHOD PRIVATE Test_FindIndexReturnsPosition
TcUnit.TEST(__POUNAME());

list.Clear();
list.AddItem(ADR(a));
list.AddItem(ADR(b));
AssertEquals_INT(Expected := 1, Actual := list.FindIndex(ADR(b)), Message := 'index of the second pointer');
AssertEquals_INT(Expected := -1, Actual := list.FindIndex(ADR(c)), Message := 'missing pointer gives -1');

TEST_FINISHED_NAMED(__POUNAME());
END_METHOD

METHOD PRIVATE Test_GetIndexReturnsPointer
TcUnit.TEST(__POUNAME());

list.Clear();
list.AddItem(ADR(a));
list.AddItem(ADR(b));
AssertTrue(Condition := list.GetIndex(1) = ADR(b), Message := 'pointer at index 1');
AssertTrue(Condition := list.GetIndex(7) = 0, Message := 'out of range gives null');

TEST_FINISHED_NAMED(__POUNAME());
END_METHOD

METHOD PRIVATE Test_RemoveIndexShiftsItems
VAR
  ok : BOOL;
END_VAR
TcUnit.TEST(__POUNAME());

list.Clear();
list.AddItem(ADR(a));
list.AddItem(ADR(b));
list.AddItem(ADR(c));
ok := list.RemoveIndex(0);
AssertTrue(Condition := ok, Message := 'remove succeeds');
AssertEquals_UDINT(Expected := 2, Actual := list.Count, Message := 'count after remove');
AssertTrue(Condition := list.GetIndex(0) = ADR(b), Message := 'second pointer shifted to the front');
AssertTrue(Condition := list.GetIndex(1) = ADR(c), Message := 'third pointer shifted down');

TEST_FINISHED_NAMED(__POUNAME());
END_METHOD

METHOD PRIVATE Test_ClearEmptiesList
TcUnit.TEST(__POUNAME());

list.Clear();
list.AddItem(ADR(a));
list.Clear();
AssertEquals_UDINT(Expected := 0, Actual := list.Count, Message := 'count after clear');
AssertFalse(Condition := list.Contains(ADR(a)), Message := 'pointers gone after clear');

TEST_FINISHED_NAMED(__POUNAME());
END_METHOD

END_FUNCTION_BLOCK

// ---- Tests/FB_LongStringList_Tests.TcPOU
FUNCTION_BLOCK FB_LongStringList_Tests EXTENDS TcUnit.FB_TestSuite
VAR
  list : FB_LongStringList;
  item : LongString;
END_VAR

Test_AddAndContains();
Test_FindIndexAndGetIndex();
Test_ContainsPartialMatchesSubstring();
Test_RemoveIndexShiftsItems();
Test_ClearEmptiesList();

METHOD PRIVATE Test_AddAndContains
TcUnit.TEST(__POUNAME());

list.Clear();
list.AddItem('alpha');
list.AddItem('beta');
AssertEquals_UDINT(Expected := 2, Actual := list.Count, Message := 'count after two adds');
AssertTrue(Condition := list.Contains('beta'), Message := 'added item found');
AssertFalse(Condition := list.Contains('gamma'), Message := 'missing item not found');

TEST_FINISHED_NAMED(__POUNAME());
END_METHOD

METHOD PRIVATE Test_FindIndexAndGetIndex
TcUnit.TEST(__POUNAME());

list.Clear();
list.AddItem('alpha');
list.AddItem('beta');
item := list.GetIndex(0);
AssertEquals_INT(Expected := 1, Actual := list.FindIndex('beta'), Message := 'index of the second item');
AssertTrue(Condition := item = 'alpha', Message := 'item at index 0');

TEST_FINISHED_NAMED(__POUNAME());
END_METHOD

METHOD PRIVATE Test_ContainsPartialMatchesSubstring
TcUnit.TEST(__POUNAME());

list.Clear();
list.AddItem('alpha');
AssertTrue(Condition := list.ContainsPartial('lph'), Message := 'substring found');
AssertFalse(Condition := list.ContainsPartial('xyz'), Message := 'missing substring not found');

TEST_FINISHED_NAMED(__POUNAME());
END_METHOD

METHOD PRIVATE Test_RemoveIndexShiftsItems
VAR
  ok : BOOL;
END_VAR
TcUnit.TEST(__POUNAME());

list.Clear();
list.AddItem('alpha');
list.AddItem('beta');
ok := list.RemoveIndex(0);
item := list.GetIndex(0);
AssertTrue(Condition := ok, Message := 'remove succeeds');
AssertEquals_UDINT(Expected := 1, Actual := list.Count, Message := 'count after remove');
AssertTrue(Condition := item = 'beta', Message := 'remaining item shifted down');

TEST_FINISHED_NAMED(__POUNAME());
END_METHOD

METHOD PRIVATE Test_ClearEmptiesList
TcUnit.TEST(__POUNAME());

list.Clear();
list.AddItem('alpha');
list.Clear();
AssertEquals_UDINT(Expected := 0, Actual := list.Count, Message := 'count after clear');

TEST_FINISHED_NAMED(__POUNAME());
END_METHOD

END_FUNCTION_BLOCK

// ---- Tests/FB_TargList_Tests.TcPOU
FUNCTION_BLOCK FB_TargList_Tests EXTENDS TcUnit.FB_TestSuite
VAR
  list : FB_TargList;
  a : INT := 1;
  b : INT := 2;
  c : INT := 3;
END_VAR

Test_AddAndContainsByValue();
Test_FindIndexReturnsPosition();
Test_GetIndexReturnsStoredArg();
Test_RemoveIndexShiftsItems();
Test_ClearEmptiesList();

METHOD PRIVATE Test_AddAndContainsByValue
TcUnit.TEST(__POUNAME());

list.Clear();
list.AddItem(F_INT(a));
list.AddItem(F_INT(b));
AssertEquals_UDINT(Expected := 2, Actual := list.Count, Message := 'count after two adds');
AssertTrue(Condition := list.Contains(F_INT(b)), Message := 'stored value found');
AssertFalse(Condition := list.Contains(F_INT(c)), Message := 'other value not found');

TEST_FINISHED_NAMED(__POUNAME());
END_METHOD

METHOD PRIVATE Test_FindIndexReturnsPosition
TcUnit.TEST(__POUNAME());

list.Clear();
list.AddItem(F_INT(a));
list.AddItem(F_INT(b));
AssertEquals_INT(Expected := 1, Actual := list.FindIndex(F_INT(b)), Message := 'index of the second value');
AssertEquals_INT(Expected := -1, Actual := list.FindIndex(F_INT(c)), Message := 'missing value gives -1');

TEST_FINISHED_NAMED(__POUNAME());
END_METHOD

METHOD PRIVATE Test_GetIndexReturnsStoredArg
VAR
  arg : T_Arg;
END_VAR
TcUnit.TEST(__POUNAME());

list.Clear();
list.AddItem(F_INT(a));
list.AddItem(F_INT(b));
arg := list.GetIndex(1);
AssertEquals_UDINT(Expected := SIZEOF(b), Actual := arg.cbLen, Message := 'length of the stored argument');
AssertTrue(Condition := arg.pData = ADR(b), Message := 'stored argument points at the variable');
AssertTrue(Condition := arg.eType = E_ArgType.ARGTYPE_INT, Message := 'type recorded');

TEST_FINISHED_NAMED(__POUNAME());
END_METHOD

METHOD PRIVATE Test_RemoveIndexShiftsItems
VAR
  ok : BOOL;
  arg : T_Arg;
END_VAR
TcUnit.TEST(__POUNAME());

list.Clear();
list.AddItem(F_INT(a));
list.AddItem(F_INT(b));
list.AddItem(F_INT(c));
ok := list.RemoveIndex(0);
arg := list.GetIndex(0);
AssertTrue(Condition := ok, Message := 'remove succeeds');
AssertEquals_UDINT(Expected := 2, Actual := list.Count, Message := 'count after remove');
AssertTrue(Condition := arg.pData = ADR(b), Message := 'second argument shifted to the front');

TEST_FINISHED_NAMED(__POUNAME());
END_METHOD

METHOD PRIVATE Test_ClearEmptiesList
TcUnit.TEST(__POUNAME());

list.Clear();
list.AddItem(F_INT(a));
list.Clear();
AssertEquals_UDINT(Expected := 0, Actual := list.Count, Message := 'count after clear');
AssertFalse(Condition := list.Contains(F_INT(a)), Message := 'values gone after clear');

TEST_FINISHED_NAMED(__POUNAME());
END_METHOD

END_FUNCTION_BLOCK

// ---- Tests/FB_Dictionary_Tests.TcPOU
FUNCTION_BLOCK FB_Dictionary_Tests EXTENDS TcUnit.FB_TestSuite
VAR
  dict : FB_Dictionary;
  a : INT := 10;
  b : INT := 20;
  c : INT := 30;
  value : T_Arg;
  key : T_MaxString;
END_VAR

Test_AddItemStoresKeyAndValue();
Test_RejectsDuplicateKey();
Test_RejectsEmptyKey();
Test_RejectsEmptyValue();
Test_TryGetReturnsValue();
Test_TryGetFailsForMissingKey();
Test_GetReturnsValue();
Test_RemoveDeletesKey();
Test_RemoveFailsForMissingKey();
Test_TryGetIndexReturnsPair();
Test_TryGetPartialKeyMatchesSubstring();
Test_ClearEmptiesDictionary();
Test_RejectsAddWhenFull();

METHOD PRIVATE Test_AddItemStoresKeyAndValue
VAR
  ok : BOOL;
  p : POINTER TO INT;
END_VAR
TcUnit.TEST(__POUNAME());

dict.Clear();
ok := dict.AddItem('a', F_INT(a));
AssertTrue(Condition := ok, Message := 'add succeeds');
AssertEquals_UDINT(Expected := 1, Actual := dict.Count, Message := 'count after one add');
AssertTrue(Condition := dict.Contains('a'), Message := 'key found');

TEST_FINISHED_NAMED(__POUNAME());
END_METHOD

METHOD PRIVATE Test_RejectsDuplicateKey
VAR
  ok : BOOL;
  p : POINTER TO INT;
END_VAR
TcUnit.TEST(__POUNAME());

dict.Clear();
dict.AddItem('a', F_INT(a));
ok := dict.AddItem('a', F_INT(b));
AssertFalse(Condition := ok, Message := 'duplicate key rejected');
AssertEquals_UDINT(Expected := 1, Actual := dict.Count, Message := 'count unchanged');

TEST_FINISHED_NAMED(__POUNAME());
END_METHOD

METHOD PRIVATE Test_RejectsEmptyKey
VAR
  ok : BOOL;
  p : POINTER TO INT;
END_VAR
TcUnit.TEST(__POUNAME());

dict.Clear();
ok := dict.AddItem('', F_INT(a));
AssertFalse(Condition := ok, Message := 'empty key rejected');
AssertEquals_UDINT(Expected := 0, Actual := dict.Count, Message := 'nothing added');

TEST_FINISHED_NAMED(__POUNAME());
END_METHOD

METHOD PRIVATE Test_RejectsEmptyValue
VAR
  ok : BOOL;
  empty : T_Arg;
END_VAR
TcUnit.TEST(__POUNAME());

dict.Clear();
ok := dict.AddItem('a', empty);
AssertFalse(Condition := ok, Message := 'zero-length value rejected');
AssertEquals_UDINT(Expected := 0, Actual := dict.Count, Message := 'nothing added');

TEST_FINISHED_NAMED(__POUNAME());
END_METHOD

METHOD PRIVATE Test_TryGetReturnsValue
VAR
  ok : BOOL;
  p : POINTER TO INT;
END_VAR
TcUnit.TEST(__POUNAME());

dict.Clear();
dict.AddItem('a', F_INT(a));
dict.AddItem('b', F_INT(b));
ok := dict.TryGet('b', value);
p := value.pData;
AssertTrue(Condition := ok, Message := 'key found');
AssertTrue(Condition := value.pData = ADR(b), Message := 'value points at the stored variable');
AssertEquals_INT(Expected := 20, Actual := p^, Message := 'value readable through the argument');

TEST_FINISHED_NAMED(__POUNAME());
END_METHOD

METHOD PRIVATE Test_TryGetFailsForMissingKey
VAR
  ok : BOOL;
  p : POINTER TO INT;
END_VAR
TcUnit.TEST(__POUNAME());

dict.Clear();
dict.AddItem('a', F_INT(a));
ok := dict.TryGet('zzz', value);
AssertFalse(Condition := ok, Message := 'missing key fails');

TEST_FINISHED_NAMED(__POUNAME());
END_METHOD

METHOD PRIVATE Test_GetReturnsValue
VAR
  ok : BOOL;
  p : POINTER TO INT;
END_VAR
TcUnit.TEST(__POUNAME());

dict.Clear();
dict.AddItem('a', F_INT(a));
value := dict.Get('a');
p := value.pData;
AssertEquals_INT(Expected := 10, Actual := p^, Message := 'Get returns the stored value');

TEST_FINISHED_NAMED(__POUNAME());
END_METHOD

METHOD PRIVATE Test_RemoveDeletesKey
VAR
  ok : BOOL;
  p : POINTER TO INT;
END_VAR
TcUnit.TEST(__POUNAME());

dict.Clear();
dict.AddItem('a', F_INT(a));
dict.AddItem('b', F_INT(b));
ok := dict.Remove('a');
AssertTrue(Condition := ok, Message := 'remove succeeds');
AssertEquals_UDINT(Expected := 1, Actual := dict.Count, Message := 'count after remove');
AssertFalse(Condition := dict.Contains('a'), Message := 'removed key gone');
AssertTrue(Condition := dict.TryGet('b', value), Message := 'other key still readable');
AssertTrue(Condition := value.pData = ADR(b), Message := 'other value intact');

TEST_FINISHED_NAMED(__POUNAME());
END_METHOD

METHOD PRIVATE Test_RemoveFailsForMissingKey
VAR
  ok : BOOL;
  p : POINTER TO INT;
END_VAR
TcUnit.TEST(__POUNAME());

dict.Clear();
dict.AddItem('a', F_INT(a));
ok := dict.Remove('zzz');
AssertFalse(Condition := ok, Message := 'missing key cannot be removed');
AssertEquals_UDINT(Expected := 1, Actual := dict.Count, Message := 'count unchanged');

TEST_FINISHED_NAMED(__POUNAME());
END_METHOD

METHOD PRIVATE Test_TryGetIndexReturnsPair
VAR
  ok : BOOL;
  p : POINTER TO INT;
END_VAR
TcUnit.TEST(__POUNAME());

dict.Clear();
dict.AddItem('a', F_INT(a));
dict.AddItem('b', F_INT(b));
ok := dict.TryGetIndex(1, key, value);
AssertTrue(Condition := ok, Message := 'index in range');
AssertEquals_STRING(Expected := 'b', Actual := key, Message := 'key at index 1');
AssertTrue(Condition := value.pData = ADR(b), Message := 'value at index 1');
AssertFalse(Condition := dict.TryGetIndex(5, key, value), Message := 'index out of range fails');

TEST_FINISHED_NAMED(__POUNAME());
END_METHOD

METHOD PRIVATE Test_TryGetPartialKeyMatchesSubstring
VAR
  ok : BOOL;
  partial : T_MaxString;
END_VAR
TcUnit.TEST(__POUNAME());

dict.Clear();
dict.AddItem('temperature', F_INT(a));
dict.AddItem('pressure', F_INT(b));
partial := 'press';
ok := dict.TryGetPartialKey(partial, value);
AssertTrue(Condition := ok, Message := 'partial key found');
AssertTrue(Condition := value.pData = ADR(b), Message := 'value of the matching key');
partial := 'flow';
AssertFalse(Condition := dict.TryGetPartialKey(partial, value), Message := 'no match fails');

TEST_FINISHED_NAMED(__POUNAME());
END_METHOD

METHOD PRIVATE Test_ClearEmptiesDictionary
TcUnit.TEST(__POUNAME());

dict.Clear();
dict.AddItem('a', F_INT(a));
dict.Clear();
AssertEquals_UDINT(Expected := 0, Actual := dict.Count, Message := 'count after clear');
AssertFalse(Condition := dict.Contains('a'), Message := 'keys gone after clear');

TEST_FINISHED_NAMED(__POUNAME());
END_METHOD

METHOD PRIVATE Test_RejectsAddWhenFull
VAR
  i : UINT;
  ok : BOOL;
END_VAR
TcUnit.TEST(__POUNAME());

dict.Clear();
FOR i := 1 TO GVL_List.LIST_SIZE DO
  dict.AddItem(CONCAT('k', TO_STRING(i)), F_INT(a));
END_FOR
ok := dict.AddItem('extra', F_INT(b));
AssertEquals_UDINT(Expected := TO_UDINT(GVL_List.LIST_SIZE), Actual := dict.Count, Message := 'dictionary holds LIST_SIZE items');
AssertFalse(Condition := ok, Message := 'add rejected when full');

TEST_FINISHED_NAMED(__POUNAME());
END_METHOD

END_FUNCTION_BLOCK

// ---- Tests/F_DictionaryValuesCrc_Tests.TcPOU
FUNCTION_BLOCK F_DictionaryValuesCrc_Tests EXTENDS TcUnit.FB_TestSuite
VAR
  dict : FB_Dictionary;
  first : INT := 1234;
  second : INT := 5678;
END_VAR

Test_EmptyDictionaryGivesZero();
Test_CrcCoversAllValues();
Test_CrcChangesWhenLaterValueChanges();

METHOD PRIVATE Test_EmptyDictionaryGivesZero
TcUnit.TEST(__POUNAME());

dict.Clear();
AssertEquals_WORD(Expected := 0, Actual := F_DictionaryValuesCrc(dict), Message := 'no values, no CRC');

TEST_FINISHED_NAMED(__POUNAME());
END_METHOD

METHOD PRIVATE Test_CrcCoversAllValues
VAR
  expected : WORD;
  actual : WORD;
END_VAR
TcUnit.TEST(__POUNAME());

// arrange
dict.Clear();
dict.AddItem('first', F_INT(first));
dict.AddItem('second', F_INT(second));
expected := F_DATA_TO_CRC16_CCITT(pData := ADR(first), cbData := SIZEOF(first), crc := 16#FFFF);
expected := F_DATA_TO_CRC16_CCITT(pData := ADR(second), cbData := SIZEOF(second), crc := expected);

// act
actual := F_DictionaryValuesCrc(dict);

// assert
AssertEquals_WORD(Expected := expected, Actual := actual, Message := 'CRC chained over every value in order');

TEST_FINISHED_NAMED(__POUNAME());
END_METHOD

METHOD PRIVATE Test_CrcChangesWhenLaterValueChanges
VAR
  before : WORD;
  after : WORD;
END_VAR
TcUnit.TEST(__POUNAME());

// arrange
dict.Clear();
dict.AddItem('first', F_INT(first));
dict.AddItem('second', F_INT(second));
before := F_DictionaryValuesCrc(dict);

// act
second := second + 1;
after := F_DictionaryValuesCrc(dict);
second := second - 1;

// assert
AssertTrue(Condition := before <> after, Message := 'a change in the second value changes the CRC');

TEST_FINISHED_NAMED(__POUNAME());
END_METHOD

END_FUNCTION_BLOCK

// ---- Tests/FB_AlphaBetaFilter_Tests.TcPOU
FUNCTION_BLOCK FB_AlphaBetaFilter_Tests EXTENDS TcUnit.FB_TestSuite

Test_UnityAlphaTracksMeasurement();
Test_HalfAlphaMovesHalfway();
Test_ZeroDeltaDoesNotDivideByZero();
Test_ConvergesToConstantInput();

METHOD PRIVATE Test_UnityAlphaTracksMeasurement
VAR
  filter : FB_AlphaBetaFilter;
END_VAR
TcUnit.TEST(__POUNAME());

filter(measurement := 10.0, deltaInSecond := 0.01, alpha := 1.0, beta := 0.0);
AssertEquals_LREAL(Expected := 10.0, Actual := filter.output, Delta := 1.0E-9, Message := 'alpha 1 passes the measurement through');

TEST_FINISHED_NAMED(__POUNAME());
END_METHOD

METHOD PRIVATE Test_HalfAlphaMovesHalfway
VAR
  filter : FB_AlphaBetaFilter;
END_VAR
TcUnit.TEST(__POUNAME());

filter(measurement := 10.0, deltaInSecond := 0.01, alpha := 0.5, beta := 0.0);
AssertEquals_LREAL(Expected := 5.0, Actual := filter.output, Delta := 1.0E-9, Message := 'first step halfway from 0');
filter(measurement := 10.0, deltaInSecond := 0.01, alpha := 0.5, beta := 0.0);
AssertEquals_LREAL(Expected := 7.5, Actual := filter.output, Delta := 1.0E-9, Message := 'second step halfway again');

TEST_FINISHED_NAMED(__POUNAME());
END_METHOD

METHOD PRIVATE Test_ZeroDeltaDoesNotDivideByZero
VAR
  filter : FB_AlphaBetaFilter;
END_VAR
TcUnit.TEST(__POUNAME());

filter(measurement := 10.0, deltaInSecond := 0.0, alpha := 0.5, beta := 0.1);
AssertEquals_LREAL(Expected := 5.0, Actual := filter.output, Delta := 1.0E-9, Message := 'velocity term dropped when delta is 0');

TEST_FINISHED_NAMED(__POUNAME());
END_METHOD

METHOD PRIVATE Test_ConvergesToConstantInput
VAR
  filter : FB_AlphaBetaFilter;
  i : INT;
END_VAR
TcUnit.TEST(__POUNAME());

FOR i := 1 TO 500 DO
  filter(measurement := 100.0, deltaInSecond := 0.01, alpha := 0.3, beta := 0.01);
END_FOR
AssertEquals_LREAL(Expected := 100.0, Actual := filter.output, Delta := 0.001, Message := 'filter settles on a constant input');

TEST_FINISHED_NAMED(__POUNAME());
END_METHOD

END_FUNCTION_BLOCK

// ---- Tests/FB_P_Control_Tests.TcPOU
FUNCTION_BLOCK FB_P_Control_Tests EXTENDS TcUnit.FB_TestSuite

Test_TermIsErrorTimesGain();
Test_NegativeErrorGivesNegativeTerm();

METHOD PRIVATE Test_TermIsErrorTimesGain
VAR
  p : FB_P_Control;
END_VAR
TcUnit.TEST(__POUNAME());

p(ProcessVariable := 4.0, Setpoint := 10.0, Kp := 2.0);
AssertEquals_LREAL(Expected := 12.0, Actual := p.Term, Delta := 1.0E-9, Message := '(10 - 4) * 2');

TEST_FINISHED_NAMED(__POUNAME());
END_METHOD

METHOD PRIVATE Test_NegativeErrorGivesNegativeTerm
VAR
  p : FB_P_Control;
END_VAR
TcUnit.TEST(__POUNAME());

p(ProcessVariable := 10.0, Setpoint := 4.0, Kp := 0.5);
AssertEquals_LREAL(Expected := -3.0, Actual := p.Term, Delta := 1.0E-9, Message := '(4 - 10) * 0.5');

TEST_FINISHED_NAMED(__POUNAME());
END_METHOD

END_FUNCTION_BLOCK

// ---- Tests/FB_I_Controller_Tests.TcPOU
FUNCTION_BLOCK FB_I_Controller_Tests EXTENDS TcUnit.FB_TestSuite

Test_IntegratesErrorOverOneCycle();
Test_AccumulatesOverCycles();
Test_ClampsAtMaximum();
Test_ClampsAtMinimum();
Test_PauseHoldsTerm();
Test_ResetClearsIntegral();
Test_ZeroGainGivesZero();
Test_UsesCycleTimeOfCallingTask();

METHOD PRIVATE Test_IntegratesErrorOverOneCycle
VAR
  i : FB_I_Controller;
  n : INT;
END_VAR
TcUnit.TEST(__POUNAME());

// the test task runs at 10 ms, so one cycle adds Ki * error * 0.01
i(ProcessVariable := 0.0, Setpoint := 1.0, Ki := 1.0, MaxIntegralComponent := 1000.0, MinIntegralComponent := -1000.0);
AssertEquals_LREAL(Expected := 0.01, Actual := i.Term, Delta := 1.0E-6, Message := 'one cycle of integration');

TEST_FINISHED_NAMED(__POUNAME());
END_METHOD

METHOD PRIVATE Test_AccumulatesOverCycles
VAR
  i : FB_I_Controller;
  n : INT;
END_VAR
TcUnit.TEST(__POUNAME());

FOR n := 1 TO 10 DO
  i(ProcessVariable := 0.0, Setpoint := 1.0, Ki := 1.0, MaxIntegralComponent := 1000.0, MinIntegralComponent := -1000.0);
END_FOR
AssertEquals_LREAL(Expected := 0.1, Actual := i.Term, Delta := 1.0E-6, Message := 'ten cycles of integration');

TEST_FINISHED_NAMED(__POUNAME());
END_METHOD

METHOD PRIVATE Test_ClampsAtMaximum
VAR
  i : FB_I_Controller;
  n : INT;
END_VAR
TcUnit.TEST(__POUNAME());

FOR n := 1 TO 10 DO
  i(ProcessVariable := 0.0, Setpoint := 1.0, Ki := 1.0, MaxIntegralComponent := 0.05, MinIntegralComponent := -1000.0);
END_FOR
AssertEquals_LREAL(Expected := 0.05, Actual := i.Term, Delta := 1.0E-9, Message := 'integral held at the maximum');

TEST_FINISHED_NAMED(__POUNAME());
END_METHOD

METHOD PRIVATE Test_ClampsAtMinimum
VAR
  i : FB_I_Controller;
  n : INT;
END_VAR
TcUnit.TEST(__POUNAME());

FOR n := 1 TO 10 DO
  i(ProcessVariable := 0.0, Setpoint := -1.0, Ki := 1.0, MaxIntegralComponent := 1000.0, MinIntegralComponent := -0.05);
END_FOR
AssertEquals_LREAL(Expected := -0.05, Actual := i.Term, Delta := 1.0E-9, Message := 'integral held at the minimum');

TEST_FINISHED_NAMED(__POUNAME());
END_METHOD

METHOD PRIVATE Test_PauseHoldsTerm
VAR
  i : FB_I_Controller;
  n : INT;
END_VAR
TcUnit.TEST(__POUNAME());

FOR n := 1 TO 5 DO
  i(ProcessVariable := 0.0, Setpoint := 1.0, Ki := 1.0, MaxIntegralComponent := 1000.0, MinIntegralComponent := -1000.0);
END_FOR
FOR n := 1 TO 5 DO
  i(ProcessVariable := 0.0, Setpoint := 1.0, Ki := 1.0, MaxIntegralComponent := 1000.0, MinIntegralComponent := -1000.0, Pause := TRUE);
END_FOR
AssertEquals_LREAL(Expected := 0.05, Actual := i.Term, Delta := 1.0E-6, Message := 'no integration while paused');

TEST_FINISHED_NAMED(__POUNAME());
END_METHOD

METHOD PRIVATE Test_ResetClearsIntegral
VAR
  i : FB_I_Controller;
  n : INT;
END_VAR
TcUnit.TEST(__POUNAME());

FOR n := 1 TO 5 DO
  i(ProcessVariable := 0.0, Setpoint := 1.0, Ki := 1.0, MaxIntegralComponent := 1000.0, MinIntegralComponent := -1000.0);
END_FOR
i(ProcessVariable := 0.0, Setpoint := 1.0, Ki := 1.0, MaxIntegralComponent := 1000.0, MinIntegralComponent := -1000.0, Reset := TRUE);
AssertEquals_LREAL(Expected := 0.01, Actual := i.Term, Delta := 1.0E-6, Message := 'reset restarts integration from zero');

TEST_FINISHED_NAMED(__POUNAME());
END_METHOD

METHOD PRIVATE Test_ZeroGainGivesZero
VAR
  i : FB_I_Controller;
  n : INT;
END_VAR
TcUnit.TEST(__POUNAME());

i(ProcessVariable := 0.0, Setpoint := 1.0, Ki := 0.0, MaxIntegralComponent := 1000.0, MinIntegralComponent := -1000.0);
AssertEquals_LREAL(Expected := 0.0, Actual := i.Term, Delta := 1.0E-9, Message := 'no gain, no term');

TEST_FINISHED_NAMED(__POUNAME());
END_METHOD

METHOD PRIVATE Test_UsesCycleTimeOfCallingTask
TcUnit.TEST(__POUNAME());

IF NOT ControllersInSlowTask.HasRunOnce THEN
  RETURN;
END_IF

AssertEquals_LREAL(Expected := 0.05, Actual := ControllersInSlowTask.IntegratorTerm, Delta := 1.0E-6, Message := 'one cycle of the 50 ms SlowTask, not the 10 ms PlcTask');

TEST_FINISHED_NAMED(__POUNAME());
END_METHOD

END_FUNCTION_BLOCK

// ---- ControllersInSlowTask.TcPOU
PROGRAM ControllersInSlowTask
VAR_OUTPUT
  HasRunOnce : BOOL;
  IntegratorTerm : LREAL;
  PiOutput : LREAL;
END_VAR
VAR
  integrator : FB_I_Controller;
  piController : FB_PI_Controller;
END_VAR

IF HasRunOnce THEN
  RETURN;
END_IF

integrator(ProcessVariable := 0.0, Setpoint := 1.0, Ki := 1.0);
piController(ProcessVariable := 0.0, Setpoint := 1.0, Kp := 0.0, IntegralConstant := 60.0, MaxLoopOutput := 100.0, MinLoopOutput := -100.0);
IntegratorTerm := integrator.Term;
PiOutput := piController.Output;
HasRunOnce := TRUE;

END_PROGRAM

// ---- Tests/FB_PI_Controller_Tests.TcPOU
FUNCTION_BLOCK FB_PI_Controller_Tests EXTENDS TcUnit.FB_TestSuite

Test_ProportionalOnlyWithBias();
Test_OutputClampedToMax();
Test_OutputClampedToMin();
Test_IntegralInRepeatsPerMinute();
Test_IntegralInRepeatsPerSecond();
Test_UsesCycleTimeOfCallingTask();

METHOD PRIVATE Test_ProportionalOnlyWithBias
VAR
  pi : FB_PI_Controller;
END_VAR
TcUnit.TEST(__POUNAME());

pi(ProcessVariable := 4.0, Setpoint := 10.0, Kp := 2.0, IntegralConstant := 0.0, MaxLoopOutput := 100.0, MinLoopOutput := -100.0, Bias := 1.0);
AssertEquals_LREAL(Expected := 13.0, Actual := pi.Output, Delta := 1.0E-9, Message := 'Kp * error + bias');

TEST_FINISHED_NAMED(__POUNAME());
END_METHOD

METHOD PRIVATE Test_OutputClampedToMax
VAR
  pi : FB_PI_Controller;
END_VAR
TcUnit.TEST(__POUNAME());

pi(ProcessVariable := 4.0, Setpoint := 10.0, Kp := 2.0, IntegralConstant := 0.0, MaxLoopOutput := 5.0, MinLoopOutput := -100.0, Bias := 0.0);
AssertEquals_LREAL(Expected := 5.0, Actual := pi.Output, Delta := 1.0E-9, Message := 'output held at the maximum');

TEST_FINISHED_NAMED(__POUNAME());
END_METHOD

METHOD PRIVATE Test_OutputClampedToMin
VAR
  pi : FB_PI_Controller;
END_VAR
TcUnit.TEST(__POUNAME());

pi(ProcessVariable := 10.0, Setpoint := 4.0, Kp := 2.0, IntegralConstant := 0.0, MaxLoopOutput := 100.0, MinLoopOutput := -5.0, Bias := 0.0);
AssertEquals_LREAL(Expected := -5.0, Actual := pi.Output, Delta := 1.0E-9, Message := 'output held at the minimum');

TEST_FINISHED_NAMED(__POUNAME());
END_METHOD

METHOD PRIVATE Test_IntegralInRepeatsPerMinute
VAR
  pi : FB_PI_Controller;
END_VAR
TcUnit.TEST(__POUNAME());

// 60 repeats per minute is 1 repeat per second: one 10 ms cycle adds error * 0.01
pi(ProcessVariable := 0.0, Setpoint := 1.0, Kp := 0.0, IntegralConstant := 60.0, RepeatsPerMinute := TRUE, MaxLoopOutput := 100.0, MinLoopOutput := -100.0, Bias := 0.0);
AssertEquals_LREAL(Expected := 0.01, Actual := pi.Output, Delta := 1.0E-6, Message := 'integral normalised from repeats per minute');

TEST_FINISHED_NAMED(__POUNAME());
END_METHOD

METHOD PRIVATE Test_IntegralInRepeatsPerSecond
VAR
  pi : FB_PI_Controller;
END_VAR
TcUnit.TEST(__POUNAME());

pi(ProcessVariable := 0.0, Setpoint := 1.0, Kp := 0.0, IntegralConstant := 1.0, RepeatsPerMinute := FALSE, MaxLoopOutput := 100.0, MinLoopOutput := -100.0, Bias := 0.0);
AssertEquals_LREAL(Expected := 0.01, Actual := pi.Output, Delta := 1.0E-6, Message := 'integral in repeats per second');

TEST_FINISHED_NAMED(__POUNAME());
END_METHOD

METHOD PRIVATE Test_UsesCycleTimeOfCallingTask
TcUnit.TEST(__POUNAME());

IF NOT ControllersInSlowTask.HasRunOnce THEN
  RETURN;
END_IF

AssertEquals_LREAL(Expected := 0.05, Actual := ControllersInSlowTask.PiOutput, Delta := 1.0E-6, Message := 'one cycle of the 50 ms SlowTask, not the 10 ms PlcTask');

TEST_FINISHED_NAMED(__POUNAME());
END_METHOD

END_FUNCTION_BLOCK

// ---- Tests/T_Task_Tests.TcPOU
FUNCTION_BLOCK T_Task_Tests EXTENDS TcUnit.FB_TestSuite
VAR
  task : T_Task;
END_VAR

Test_NameIsPlcTask();
Test_CycleTimeMatchesConfiguredTask();
Test_CycleCountAdvances();
Test_DistributedClockUnitsAgree();
Test_DateTimeStringFormat();
Test_DateStringIsDateOnly();
Test_TimeStringIsTimeOnly();
Test_DateTimeFromDcIsCurrent();
Test_SetToThisTaskSelectsCurrentTask();

METHOD PRIVATE Test_NameIsPlcTask
TcUnit.TEST(__POUNAME());

AssertEquals_STRING(Expected := 'PlcTask', Actual := RIGHT(task.Name, 7), Message := 'task name read from _TaskInfo ends with the task name');
AssertTrue(Condition := LEN(task.Name) >= 7, Message := 'task name is not empty');

TEST_FINISHED_NAMED(__POUNAME());
END_METHOD

METHOD PRIVATE Test_CycleTimeMatchesConfiguredTask
TcUnit.TEST(__POUNAME());

AssertEquals_LREAL(Expected := 10.0, Actual := task.CycleTimeInMs, Delta := 1.0E-6, Message := 'PlcTask runs every 10 ms');
AssertEquals_LREAL(Expected := 0.01, Actual := task.CycleTimeInSecs, Delta := 1.0E-9, Message := 'cycle time in seconds');
AssertEquals_LREAL(Expected := 100.0, Actual := task.CyclesPerSecond, Delta := 1.0E-6, Message := 'cycles per second');

TEST_FINISHED_NAMED(__POUNAME());
END_METHOD

METHOD PRIVATE Test_CycleCountAdvances
TcUnit.TEST(__POUNAME());

AssertTrue(Condition := task.CycleCount > 0, Message := 'cycle count read from _TaskInfo');

TEST_FINISHED_NAMED(__POUNAME());
END_METHOD

METHOD PRIVATE Test_DistributedClockUnitsAgree
VAR
  ns : LINT;
  ms : LINT;
END_VAR
TcUnit.TEST(__POUNAME());

ns := task.DistributedClockTimeInNs;
ms := task.DistributedClockTimeInMs;
AssertEquals_LINT(Expected := ns / 1000000, Actual := ms, Message := 'milliseconds derived from nanoseconds');
AssertEquals_LINT(Expected := ms / 1000, Actual := task.DistributedClockTimeInSecs, Message := 'seconds derived from milliseconds');
AssertTrue(Condition := ns > 0, Message := 'distributed clock is running');

TEST_FINISHED_NAMED(__POUNAME());
END_METHOD

METHOD PRIVATE Test_DateTimeStringFormat
VAR
  text : STRING;
END_VAR
TcUnit.TEST(__POUNAME());

// yyyy-mm-dd_hh-mm-ss
text := task.DateTimeString;
AssertEquals_INT(Expected := 19, Actual := LEN(text), Message := 'length of yyyy-mm-dd_hh-mm-ss');
AssertEquals_BYTE(Expected := 45, Actual := text[4], Message := 'dash after the year');
AssertEquals_BYTE(Expected := 45, Actual := text[7], Message := 'dash after the month');
AssertEquals_BYTE(Expected := 95, Actual := text[10], Message := 'underscore between date and time');
AssertEquals_BYTE(Expected := 45, Actual := text[13], Message := 'dash after the hour');
AssertEquals_BYTE(Expected := 45, Actual := text[16], Message := 'dash after the minute');

TEST_FINISHED_NAMED(__POUNAME());
END_METHOD

METHOD PRIVATE Test_DateStringIsDateOnly
VAR
  text : STRING;
END_VAR
TcUnit.TEST(__POUNAME());

text := task.DateString;
AssertEquals_INT(Expected := 10, Actual := LEN(text), Message := 'length of yyyy-mm-dd');
AssertEquals_STRING(Expected := LEFT(task.DateTimeString, 10), Actual := text, Message := 'date part of the date-time string');

TEST_FINISHED_NAMED(__POUNAME());
END_METHOD

METHOD PRIVATE Test_TimeStringIsTimeOnly
VAR
  text : STRING;
END_VAR
TcUnit.TEST(__POUNAME());

text := task.TimeString;
AssertEquals_INT(Expected := 8, Actual := LEN(text), Message := 'length of hh-mm-ss');
AssertEquals_STRING(Expected := RIGHT(task.DateTimeString, 8), Actual := text, Message := 'time part of the date-time string');

TEST_FINISHED_NAMED(__POUNAME());
END_METHOD

METHOD PRIVATE Test_DateTimeFromDcIsCurrent
TcUnit.TEST(__POUNAME());

AssertTrue(Condition := task.DateTimeFromDc > DT#2026-01-01-00:00:00, Message := 'distributed clock converts to a current date');

TEST_FINISHED_NAMED(__POUNAME());
END_METHOD

METHOD PRIVATE Test_SetToThisTaskSelectsCurrentTask
TcUnit.TEST(__POUNAME());

task.Index := 7;
task.SetToThisTask();
AssertEquals_BYTE(Expected := 1, Actual := task.Index, Message := 'PlcTask is the first task of the test runner');

TEST_FINISHED_NAMED(__POUNAME());
END_METHOD

END_FUNCTION_BLOCK

// ---- Tests/T_NamedBase_Tests.TcPOU
FUNCTION_BLOCK T_NamedBase_Tests EXTENDS TcUnit.FB_TestSuite
VAR
  named : T_NamedBase;
  mock : T_MockExternalLogger;
END_VAR

Test_ObjectNameIsDeclaredName();
Test_InstanceNameStartsAtProgram();
Test_LogInfoPrefixesInstanceName();

METHOD PRIVATE Test_ObjectNameIsDeclaredName
TcUnit.TEST(__POUNAME());

AssertEquals_STRING(Expected := 'named', Actual := named.ObjectName, Message := 'object name is the last segment of the instance path');

TEST_FINISHED_NAMED(__POUNAME());
END_METHOD

METHOD PRIVATE Test_InstanceNameStartsAtProgram
VAR
  name : T_MaxString;
END_VAR
TcUnit.TEST(__POUNAME());

name := named.InstanceName;
AssertEquals_STRING(Expected := 'MAIN.suiteNamedBase.named', Actual := name, Message := 'instance name starts at the program, project name removed');

TEST_FINISHED_NAMED(__POUNAME());
END_METHOD

METHOD PRIVATE Test_LogInfoPrefixesInstanceName
TcUnit.TEST(__POUNAME());

// arrange
LogConfig.ExternalLogger := mock;
LogConfig.LogLevel := E_LogSeverity.Debug;
mock.Reset();

// act
named.LogInfo('hello');

// assert
AssertEquals_STRING(Expected := CONCAT(named.InstanceName, ': hello'), Actual := mock.LastMessage, Message := 'message carries the instance name');
AssertTrue(Condition := mock.LastSeverity = E_LogSeverity.Info, Message := 'logged as info');

// cleanup
LogConfig.LogLevel := E_LogSeverity.None;
LogConfig.ExternalLogger := 0;

TEST_FINISHED_NAMED(__POUNAME());
END_METHOD

END_FUNCTION_BLOCK

// ---- Mocks/T_MockExternalLogger.TcPOU
// Test double for I_ExternalLogger: records the last message and severity.
FUNCTION_BLOCK T_MockExternalLogger IMPLEMENTS I_ExternalLogger
VAR
  _lastMessage : T_MaxString;
  _lastSeverity : E_LogSeverity;
  _callCount : UDINT;
END_VAR

METHOD AddToLog
VAR_IN_OUT
  Message : T_MaxString;
END_VAR
VAR_INPUT
  LogSeverity : E_LogSeverity;
END_VAR
_lastMessage := Message;
_lastSeverity := LogSeverity;
_callCount := _callCount + 1;
END_METHOD

METHOD Reset
_lastMessage := '';
_lastSeverity := E_LogSeverity.None;
_callCount := 0;
END_METHOD

PROPERTY CallCount : UDINT
GET
CallCount := _callCount;
END_GET
END_PROPERTY

PROPERTY LastMessage : T_MaxString
GET
LastMessage := _lastMessage;
END_GET
END_PROPERTY

PROPERTY LastSeverity : E_LogSeverity
GET
LastSeverity := _lastSeverity;
END_GET
END_PROPERTY

END_FUNCTION_BLOCK

// ---- Tests/Logger_Tests.TcPOU
FUNCTION_BLOCK Logger_Tests EXTENDS TcUnit.FB_TestSuite
VAR
  mock : T_MockExternalLogger;
  risingEdge : FB_LogOnEdge;
  fallingEdge : FB_LogOnEdge;
  badSeverity : FB_LogOnEdge;
  infoEdge : FB_LogInfoEdge;
  warningEdge : FB_LogWarningEdge;
  errorEdge : FB_LogErrorEdge;
END_VAR

Test_InfoLoggedAtDebugLevel();
Test_DebugMessageIsPrefixed();
Test_WarningFilteredBelowErrorLevel();
Test_ErrorPassesErrorLevel();
Test_NoneLevelSilencesEverything();
Test_SeverityToString();
Test_LogOnEdgeFiresOnRisingEdge();
Test_LogOnEdgeFiresOnFallingEdge();
Test_LogOnEdgeReportsUnsupportedSeverity();
Test_TypedEdgeWrappersUseTheirSeverity();

METHOD PRIVATE Test_InfoLoggedAtDebugLevel
VAR
  result : STRING;
END_VAR
TcUnit.TEST(__POUNAME());

UseMockAtLevel(E_LogSeverity.Debug);
result := F_LogInfo('hello');
AssertEquals_STRING(Expected := 'hello', Actual := result, Message := 'logged message returned');
AssertEquals_UDINT(Expected := 1, Actual := mock.CallCount, Message := 'external logger called once');
AssertEquals_STRING(Expected := 'hello', Actual := mock.LastMessage, Message := 'message passed on');
AssertTrue(Condition := mock.LastSeverity = E_LogSeverity.Info, Message := 'severity is info');
RestoreLogConfig();

TEST_FINISHED_NAMED(__POUNAME());
END_METHOD

METHOD PRIVATE Test_DebugMessageIsPrefixed
TcUnit.TEST(__POUNAME());

UseMockAtLevel(E_LogSeverity.Debug);
F_LogDebug('x');
AssertEquals_STRING(Expected := 'DEBUG x', Actual := mock.LastMessage, Message := 'debug messages carry a DEBUG prefix');
AssertTrue(Condition := mock.LastSeverity = E_LogSeverity.Debug, Message := 'severity is debug');
RestoreLogConfig();

TEST_FINISHED_NAMED(__POUNAME());
END_METHOD

METHOD PRIVATE Test_WarningFilteredBelowErrorLevel
VAR
  result : STRING;
END_VAR
TcUnit.TEST(__POUNAME());

UseMockAtLevel(E_LogSeverity.Error);
result := F_LogWarning('w');
AssertEquals_STRING(Expected := '', Actual := result, Message := 'filtered message returns empty');
AssertEquals_UDINT(Expected := 0, Actual := mock.CallCount, Message := 'external logger not called');
RestoreLogConfig();

TEST_FINISHED_NAMED(__POUNAME());
END_METHOD

METHOD PRIVATE Test_ErrorPassesErrorLevel
TcUnit.TEST(__POUNAME());

UseMockAtLevel(E_LogSeverity.Error);
F_LogError('e');
AssertEquals_UDINT(Expected := 1, Actual := mock.CallCount, Message := 'external logger called');
AssertTrue(Condition := mock.LastSeverity = E_LogSeverity.Error, Message := 'severity is error');
RestoreLogConfig();

TEST_FINISHED_NAMED(__POUNAME());
END_METHOD

METHOD PRIVATE Test_NoneLevelSilencesEverything
VAR
  result : STRING;
END_VAR
TcUnit.TEST(__POUNAME());

UseMockAtLevel(E_LogSeverity.None);
result := F_LogError('e');
AssertEquals_STRING(Expected := '', Actual := result, Message := 'nothing logged at level None');
AssertEquals_UDINT(Expected := 0, Actual := mock.CallCount, Message := 'external logger not called');
RestoreLogConfig();

TEST_FINISHED_NAMED(__POUNAME());
END_METHOD

METHOD PRIVATE Test_SeverityToString
TcUnit.TEST(__POUNAME());

AssertEquals_STRING(Expected := 'Info', Actual := TO_STRING(E_LogSeverity.Info), Message := 'info name');
AssertEquals_STRING(Expected := 'Warning', Actual := TO_STRING(E_LogSeverity.Warning), Message := 'warning name');
AssertEquals_STRING(Expected := 'Error', Actual := TO_STRING(E_LogSeverity.Error), Message := 'error name');

TEST_FINISHED_NAMED(__POUNAME());
END_METHOD

METHOD PRIVATE Test_LogOnEdgeFiresOnRisingEdge
TcUnit.TEST(__POUNAME());

UseMockAtLevel(E_LogSeverity.Debug);
risingEdge(Event := FALSE, Message := 'rise', LogSeverity := E_LogSeverity.Info);
risingEdge(Event := TRUE, Message := 'rise', LogSeverity := E_LogSeverity.Info);
AssertTrue(Condition := risingEdge.Q, Message := 'Q on the rising edge');
AssertEquals_UDINT(Expected := 1, Actual := mock.CallCount, Message := 'logged once');
AssertEquals_STRING(Expected := 'rise', Actual := mock.LastMessage, Message := 'message logged');
risingEdge(Event := TRUE, Message := 'rise', LogSeverity := E_LogSeverity.Info);
AssertFalse(Condition := risingEdge.Q, Message := 'Q clears while the event stays set');
AssertEquals_UDINT(Expected := 1, Actual := mock.CallCount, Message := 'not logged again');
RestoreLogConfig();

TEST_FINISHED_NAMED(__POUNAME());
END_METHOD

METHOD PRIVATE Test_LogOnEdgeFiresOnFallingEdge
TcUnit.TEST(__POUNAME());

UseMockAtLevel(E_LogSeverity.Debug);
fallingEdge(Event := TRUE, Message := 'fall', LogSeverity := E_LogSeverity.Warning, EventFallingEdge := TRUE);
AssertEquals_UDINT(Expected := 0, Actual := mock.CallCount, Message := 'rising edge ignored in falling mode');
fallingEdge(Event := FALSE, Message := 'fall', LogSeverity := E_LogSeverity.Warning, EventFallingEdge := TRUE);
AssertTrue(Condition := fallingEdge.Q, Message := 'Q on the falling edge');
AssertEquals_UDINT(Expected := 1, Actual := mock.CallCount, Message := 'logged once');
AssertTrue(Condition := mock.LastSeverity = E_LogSeverity.Warning, Message := 'severity passed on');
RestoreLogConfig();

TEST_FINISHED_NAMED(__POUNAME());
END_METHOD

METHOD PRIVATE Test_LogOnEdgeReportsUnsupportedSeverity
TcUnit.TEST(__POUNAME());

UseMockAtLevel(E_LogSeverity.Debug);
badSeverity(Event := FALSE, Message := 'odd', LogSeverity := E_LogSeverity.Debug);
badSeverity(Event := TRUE, Message := 'odd', LogSeverity := E_LogSeverity.Debug);
AssertTrue(Condition := mock.LastSeverity = E_LogSeverity.Error, Message := 'an unsupported severity is reported as an error');
AssertTrue(Condition := FIND(mock.LastMessage, 'odd') > 0, Message := 'the original message is included');
RestoreLogConfig();

TEST_FINISHED_NAMED(__POUNAME());
END_METHOD

METHOD PRIVATE Test_TypedEdgeWrappersUseTheirSeverity
TcUnit.TEST(__POUNAME());

UseMockAtLevel(E_LogSeverity.Debug);
infoEdge(Event := FALSE, Message := 'i');
infoEdge(Event := TRUE, Message := 'i');
AssertTrue(Condition := infoEdge.Q, Message := 'info edge Q');
AssertTrue(Condition := mock.LastSeverity = E_LogSeverity.Info, Message := 'info edge logs info');
warningEdge(Event := FALSE, Message := 'w');
warningEdge(Event := TRUE, Message := 'w');
AssertTrue(Condition := warningEdge.Q, Message := 'warning edge Q');
AssertTrue(Condition := mock.LastSeverity = E_LogSeverity.Warning, Message := 'warning edge logs warning');
errorEdge(Event := FALSE, Message := 'e');
errorEdge(Event := TRUE, Message := 'e');
AssertTrue(Condition := errorEdge.Q, Message := 'error edge Q');
AssertTrue(Condition := mock.LastSeverity = E_LogSeverity.Error, Message := 'error edge logs error');
AssertEquals_UDINT(Expected := 3, Actual := mock.CallCount, Message := 'one log per edge');
RestoreLogConfig();

TEST_FINISHED_NAMED(__POUNAME());
END_METHOD

// Test helper: route the library logger to the mock at the given level.
METHOD PRIVATE UseMockAtLevel
VAR_INPUT
  level : E_LogSeverity;
END_VAR
LogConfig.ExternalLogger := mock;
LogConfig.LogLevel := level;
mock.Reset();
END_METHOD

// Test helper: put the library logger back to its defaults.
METHOD PRIVATE RestoreLogConfig
LogConfig.LogLevel := E_LogSeverity.None;
LogConfig.ExternalLogger := 0;
END_METHOD

END_FUNCTION_BLOCK

// ---- Tests/FB_Assert_Tests.TcPOU
FUNCTION_BLOCK FB_Assert_Tests EXTENDS TcUnit.FB_TestSuite
VAR
  assert : FB_Assert;
END_VAR

Test_IsTrue();
Test_IsFalse();
Test_FloatsAreEqualWithinPrecision();
Test_FloatsAreDifferentOutsidePrecision();

METHOD PRIVATE Test_IsTrue
TcUnit.TEST(__POUNAME());

AssertTrue(Condition := assert.IsTrue(TRUE, 'x'), Message := 'TRUE passes IsTrue');
AssertFalse(Condition := assert.IsTrue(FALSE, 'x'), Message := 'FALSE fails IsTrue');

TEST_FINISHED_NAMED(__POUNAME());
END_METHOD

METHOD PRIVATE Test_IsFalse
TcUnit.TEST(__POUNAME());

AssertTrue(Condition := assert.IsFalse(FALSE, 'x'), Message := 'FALSE passes IsFalse');
AssertFalse(Condition := assert.IsFalse(TRUE, 'x'), Message := 'TRUE fails IsFalse');

TEST_FINISHED_NAMED(__POUNAME());
END_METHOD

METHOD PRIVATE Test_FloatsAreEqualWithinPrecision
TcUnit.TEST(__POUNAME());

AssertTrue(Condition := assert.FloatsAreEqual(1.0, 1.0005, 0.001, 'x'), Message := 'within precision');
AssertFalse(Condition := assert.FloatsAreEqual(1.0, 1.1, 0.001, 'x'), Message := 'outside precision');

TEST_FINISHED_NAMED(__POUNAME());
END_METHOD

METHOD PRIVATE Test_FloatsAreDifferentOutsidePrecision
TcUnit.TEST(__POUNAME());

AssertTrue(Condition := assert.FloatsAreDifferent(1.0, 1.1, 0.001, 'x'), Message := 'outside precision');
AssertFalse(Condition := assert.FloatsAreDifferent(1.0, 1.0005, 0.001, 'x'), Message := 'within precision');

TEST_FINISHED_NAMED(__POUNAME());
END_METHOD

END_FUNCTION_BLOCK

// ---- Tests/F_GetKL306xState_Tests.TcPOU
FUNCTION_BLOCK F_GetKL306xState_Tests EXTENDS TcUnit.FB_TestSuite

Test_Limit1BitsDecode();
Test_Limit2BitsDecode();
Test_RangeAndErrorFlagsPassThrough();

METHOD PRIVATE Test_Limit1BitsDecode
VAR
  status : stKL306x_ChannelStatus;
  isEqual, isGreater, isLess, notEnabled : BOOL;
END_VAR
TcUnit.TEST(__POUNAME());

status.Limit1Bit_1 := TRUE; status.Limit1Bit_0 := TRUE;
F_GetKL306xState(KL306xState := status, ProcessData_EQ_Limit1 => isEqual, ProcessData_GT_Limit1 => isGreater, ProcessData_LT_Limit1 => isLess, Limit1NotEnabled => notEnabled);
AssertTrue(Condition := isEqual AND NOT isGreater AND NOT isLess AND NOT notEnabled, Message := '11 = equal to limit 1');

status.Limit1Bit_1 := TRUE; status.Limit1Bit_0 := FALSE;
F_GetKL306xState(KL306xState := status, ProcessData_EQ_Limit1 => isEqual, ProcessData_GT_Limit1 => isGreater, ProcessData_LT_Limit1 => isLess, Limit1NotEnabled => notEnabled);
AssertTrue(Condition := isGreater AND NOT isEqual AND NOT isLess AND NOT notEnabled, Message := '10 = greater than limit 1');

status.Limit1Bit_1 := FALSE; status.Limit1Bit_0 := TRUE;
F_GetKL306xState(KL306xState := status, ProcessData_EQ_Limit1 => isEqual, ProcessData_GT_Limit1 => isGreater, ProcessData_LT_Limit1 => isLess, Limit1NotEnabled => notEnabled);
AssertTrue(Condition := isLess AND NOT isEqual AND NOT isGreater AND NOT notEnabled, Message := '01 = less than limit 1');

status.Limit1Bit_1 := FALSE; status.Limit1Bit_0 := FALSE;
F_GetKL306xState(KL306xState := status, ProcessData_EQ_Limit1 => isEqual, ProcessData_GT_Limit1 => isGreater, ProcessData_LT_Limit1 => isLess, Limit1NotEnabled => notEnabled);
AssertTrue(Condition := notEnabled AND NOT isEqual AND NOT isGreater AND NOT isLess, Message := '00 = limit 1 not enabled');

TEST_FINISHED_NAMED(__POUNAME());
END_METHOD

METHOD PRIVATE Test_Limit2BitsDecode
VAR
  status : stKL306x_ChannelStatus;
  isEqual, isGreater, isLess, notEnabled : BOOL;
END_VAR
TcUnit.TEST(__POUNAME());

status.Limit2Bit_1 := TRUE; status.Limit2Bit_0 := TRUE;
F_GetKL306xState(KL306xState := status, ProcessData_EQ_Limit2 => isEqual, ProcessData_GT_Limit2 => isGreater, ProcessData_LT_Limit2 => isLess, Limit2NotEnabled => notEnabled);
AssertTrue(Condition := isEqual AND NOT isGreater AND NOT isLess AND NOT notEnabled, Message := '11 = equal to limit 2');

status.Limit2Bit_1 := TRUE; status.Limit2Bit_0 := FALSE;
F_GetKL306xState(KL306xState := status, ProcessData_EQ_Limit2 => isEqual, ProcessData_GT_Limit2 => isGreater, ProcessData_LT_Limit2 => isLess, Limit2NotEnabled => notEnabled);
AssertTrue(Condition := isGreater AND NOT isEqual AND NOT isLess AND NOT notEnabled, Message := '10 = greater than limit 2');

status.Limit2Bit_1 := FALSE; status.Limit2Bit_0 := TRUE;
F_GetKL306xState(KL306xState := status, ProcessData_EQ_Limit2 => isEqual, ProcessData_GT_Limit2 => isGreater, ProcessData_LT_Limit2 => isLess, Limit2NotEnabled => notEnabled);
AssertTrue(Condition := isLess AND NOT isEqual AND NOT isGreater AND NOT notEnabled, Message := '01 = less than limit 2');

status.Limit2Bit_1 := FALSE; status.Limit2Bit_0 := FALSE;
F_GetKL306xState(KL306xState := status, ProcessData_EQ_Limit2 => isEqual, ProcessData_GT_Limit2 => isGreater, ProcessData_LT_Limit2 => isLess, Limit2NotEnabled => notEnabled);
AssertTrue(Condition := notEnabled AND NOT isEqual AND NOT isGreater AND NOT isLess, Message := '00 = limit 2 not enabled');

TEST_FINISHED_NAMED(__POUNAME());
END_METHOD

METHOD PRIVATE Test_RangeAndErrorFlagsPassThrough
VAR
  status : stKL306x_ChannelStatus;
  under, over, err : BOOL;
END_VAR
TcUnit.TEST(__POUNAME());

status.Underrange := TRUE; status.Overrange := FALSE; status.Error := TRUE;
F_GetKL306xState(KL306xState := status, Underrange => under, Overrange => over, Error => err);
AssertTrue(Condition := under, Message := 'underrange passed through');
AssertFalse(Condition := over, Message := 'overrange passed through');
AssertTrue(Condition := err, Message := 'error passed through');

TEST_FINISHED_NAMED(__POUNAME());
END_METHOD

END_FUNCTION_BLOCK

// ---- Tests/ProjectInformation_Tests.TcPOU
FUNCTION_BLOCK ProjectInformation_Tests EXTENDS TcUnit.FB_TestSuite

Test_VersionIsFourPointTwo();
Test_TitleAndCompany();

METHOD PRIVATE Test_VersionIsFourPointTwo
VAR
  version : ST_LibVersion;
END_VAR
TcUnit.TEST(__POUNAME());

version := F_GetVersion();
AssertEquals_STRING(Expected := '4.2.0.0', Actual := version.sVersion, Message := 'library version string');
AssertEquals_UINT(Expected := 4, Actual := version.iMajor, Message := 'major version');
AssertEquals_UINT(Expected := 2, Actual := version.iMinor, Message := 'minor version');

TEST_FINISHED_NAMED(__POUNAME());
END_METHOD

METHOD PRIVATE Test_TitleAndCompany
TcUnit.TEST(__POUNAME());

AssertEquals_WSTRING(Expected := "Intecre.Utilities", Actual := F_GetTitle(), Message := 'library title');
AssertEquals_WSTRING(Expected := "Intecre Ltd", Actual := F_GetCompany(), Message := 'library company');

TEST_FINISHED_NAMED(__POUNAME());
END_METHOD

END_FUNCTION_BLOCK

// ---- Tests/F_TargToString_Tests.TcPOU
FUNCTION_BLOCK F_TargToString_Tests EXTENDS TcUnit.FB_TestSuite
VAR
  i : INT := 42;
  d : DINT := -7;
  lr : LREAL := 1.5;
  text : T_MaxString := 'hi';
  b : BOOL := TRUE;
  w : WORD := 16#FFFF;
  li : LINT := 5;
END_VAR

Test_IntToString();
Test_DintToString();
Test_LrealToString();
Test_StringToString();
Test_BoolToString();
Test_WordToString();
Test_UnsupportedTypeGivesEmpty();

METHOD PRIVATE Test_IntToString
TcUnit.TEST(__POUNAME());

AssertEquals_STRING(Expected := '42', Actual := F_TargToString(F_INT(i)), Message := 'INT formatted');

TEST_FINISHED_NAMED(__POUNAME());
END_METHOD

METHOD PRIVATE Test_DintToString
TcUnit.TEST(__POUNAME());

AssertEquals_STRING(Expected := '-7', Actual := F_TargToString(F_DINT(d)), Message := 'DINT formatted');

TEST_FINISHED_NAMED(__POUNAME());
END_METHOD

METHOD PRIVATE Test_LrealToString
TcUnit.TEST(__POUNAME());

AssertEquals_STRING(Expected := '1.5', Actual := F_TargToString(F_LREAL(lr)), Message := 'LREAL formatted');

TEST_FINISHED_NAMED(__POUNAME());
END_METHOD

METHOD PRIVATE Test_StringToString
TcUnit.TEST(__POUNAME());

AssertEquals_STRING(Expected := 'hi', Actual := F_TargToString(F_STRING(text)), Message := 'STRING passed through');

TEST_FINISHED_NAMED(__POUNAME());
END_METHOD

METHOD PRIVATE Test_BoolToString
TcUnit.TEST(__POUNAME());

AssertEquals_STRING(Expected := 'TRUE', Actual := F_TargToString(F_BOOL(b)), Message := 'BOOL formatted');

TEST_FINISHED_NAMED(__POUNAME());
END_METHOD

METHOD PRIVATE Test_WordToString
TcUnit.TEST(__POUNAME());

AssertEquals_STRING(Expected := '65535', Actual := F_TargToString(F_WORD(w)), Message := 'WORD formatted');

TEST_FINISHED_NAMED(__POUNAME());
END_METHOD

METHOD PRIVATE Test_UnsupportedTypeGivesEmpty
TcUnit.TEST(__POUNAME());

AssertEquals_STRING(Expected := '', Actual := F_TargToString(F_LINT(li)), Message := 'LINT is not handled and gives an empty string');

TEST_FINISHED_NAMED(__POUNAME());
END_METHOD

END_FUNCTION_BLOCK

// ---- Tests/F_StringToTarg_Tests.TcPOU
FUNCTION_BLOCK F_StringToTarg_Tests EXTENDS TcUnit.FB_TestSuite
VAR
  i : INT;
  d : DINT;
  lr : LREAL;
  text : T_MaxString;
  b : BOOL;
  li : LINT;
  targ : T_Arg;
END_VAR

Test_WritesInt();
Test_WritesDint();
Test_WritesLreal();
Test_WritesString();
Test_WritesBool();
Test_UnsupportedTypeLeavesValue();

METHOD PRIVATE Test_WritesInt
TcUnit.TEST(__POUNAME());

i := 0;
targ := F_INT(i);
F_StringToTarg('123', targ);
AssertEquals_INT(Expected := 123, Actual := i, Message := 'INT written through the argument');

TEST_FINISHED_NAMED(__POUNAME());
END_METHOD

METHOD PRIVATE Test_WritesDint
TcUnit.TEST(__POUNAME());

d := 0;
targ := F_DINT(d);
F_StringToTarg('-99', targ);
AssertEquals_DINT(Expected := -99, Actual := d, Message := 'DINT written through the argument');

TEST_FINISHED_NAMED(__POUNAME());
END_METHOD

METHOD PRIVATE Test_WritesLreal
TcUnit.TEST(__POUNAME());

lr := 0.0;
targ := F_LREAL(lr);
F_StringToTarg('2.5', targ);
AssertEquals_LREAL(Expected := 2.5, Actual := lr, Delta := 1.0E-9, Message := 'LREAL written through the argument');

TEST_FINISHED_NAMED(__POUNAME());
END_METHOD

METHOD PRIVATE Test_WritesString
TcUnit.TEST(__POUNAME());

text := '';
targ := F_STRING(text);
F_StringToTarg('abc', targ);
AssertEquals_STRING(Expected := 'abc', Actual := text, Message := 'STRING written through the argument');

TEST_FINISHED_NAMED(__POUNAME());
END_METHOD

METHOD PRIVATE Test_WritesBool
TcUnit.TEST(__POUNAME());

b := FALSE;
targ := F_BOOL(b);
F_StringToTarg('TRUE', targ);
AssertTrue(Condition := b, Message := 'BOOL written through the argument');
F_StringToTarg('FALSE', targ);
AssertFalse(Condition := b, Message := 'BOOL cleared through the argument');

TEST_FINISHED_NAMED(__POUNAME());
END_METHOD

METHOD PRIVATE Test_UnsupportedTypeLeavesValue
TcUnit.TEST(__POUNAME());

li := 5;
targ := F_LINT(li);
F_StringToTarg('9', targ);
AssertEquals_LINT(Expected := 5, Actual := li, Message := 'LINT is not handled and stays unchanged');

TEST_FINISHED_NAMED(__POUNAME());
END_METHOD

END_FUNCTION_BLOCK

// ---- Tests/F_GetAmsNetId_Tests.TcPOU
FUNCTION_BLOCK F_GetAmsNetId_Tests EXTENDS TcUnit.FB_TestSuite

Test_ZeroArrayMeansLocal();
Test_FormatsNonZeroArray();

METHOD PRIVATE Test_ZeroArrayMeansLocal
VAR
  arr : T_AmsNetIdArr;
END_VAR
TcUnit.TEST(__POUNAME());

AssertEquals_STRING(Expected := '', Actual := F_GetAmsNetId(arr), Message := 'all-zero NetId maps to the local (empty) NetId');

TEST_FINISHED_NAMED(__POUNAME());
END_METHOD

METHOD PRIVATE Test_FormatsNonZeroArray
VAR
  arr : T_AmsNetIdArr;
END_VAR
TcUnit.TEST(__POUNAME());

arr[0] := 5; arr[1] := 6; arr[2] := 7; arr[3] := 8; arr[4] := 1; arr[5] := 1;
AssertEquals_STRING(Expected := '5.6.7.8.1.1', Actual := F_GetAmsNetId(arr), Message := 'NetId formatted as dotted text');

TEST_FINISHED_NAMED(__POUNAME());
END_METHOD

END_FUNCTION_BLOCK

// ---- Tests/T_Timer_Tests.TcPOU
// Timed tests: each test is a small state machine driven every cycle.
FUNCTION_BLOCK T_Timer_Tests EXTENDS TcUnit.FB_TestSuite
VAR
  timer : T_Timer;
  pulseTimer : T_Timer;
  periodTimer : T_Timer;
END_VAR

Test_QOnAndQOffFollowThePeriod();
Test_PulseTrainTogglesEachHalfPeriod();
Test_SetPeriodReadsBackWithMinimumOfOneMs();

METHOD PRIVATE Test_QOnAndQOffFollowThePeriod
VAR_INST
  state : INT := 10;
  wait : TON;
END_VAR
TcUnit.TEST(__POUNAME());

wait();

CASE state OF

  10:

    // arrange
    timer.SetPeriod := T#50MS;
    timer.Signal := TRUE;

    // assert: nothing has elapsed yet
    AssertFalse(Condition := timer.Q_On, Message := 'Q_On is not set as soon as the signal arrives');
    AssertTrue(Condition := timer.ElapsedTimeInMs < 20, Message := 'elapsed time starts near zero');
    state := 20;
    wait(IN := TRUE, PT := T#150MS);

  20:

    IF NOT wait.Q THEN
      RETURN;
    END_IF
    wait(IN := FALSE);

    // assert: period elapsed with the signal on
    AssertTrue(Condition := timer.Q_On, Message := 'Q_On after the period has elapsed');
    AssertFalse(Condition := timer.Q_Off, Message := 'Q_Off stays clear while the signal is on');
    AssertTrue(Condition := (timer.ElapsedTimeInMs >= 100) AND (timer.ElapsedTimeInMs < 400), Message := 'elapsed time tracks the wait');
    AssertTrue(Condition := timer.ElapsedTime >= T#100MS, Message := 'elapsed time as TIME');

    // act: drop the signal
    timer.Signal := FALSE;
    AssertEquals_LINT(Expected := 0, Actual := timer.ElapsedTimeInMs, Message := 'elapsed time reads zero once the signal is off');
    AssertFalse(Condition := timer.Q_On, Message := 'Q_On clears with the signal');
    AssertFalse(Condition := timer.Q_Off, Message := 'Q_Off needs the period to elapse first');
    state := 30;
    wait(IN := TRUE, PT := T#150MS);

  30:

    IF NOT wait.Q THEN
      RETURN;
    END_IF
    wait(IN := FALSE);

    // assert: period elapsed with the signal off
    AssertTrue(Condition := timer.Q_Off, Message := 'Q_Off after the period has elapsed with the signal off');
    AssertFalse(Condition := timer.Q_On, Message := 'Q_On stays clear while the signal is off');
    TEST_FINISHED_NAMED(__POUNAME());
    state := 40;

  40:
    ; // finished

END_CASE
END_METHOD

METHOD PRIVATE Test_PulseTrainTogglesEachHalfPeriod
VAR_INST
  state : INT := 10;
  wait : TON;
END_VAR
TcUnit.TEST(__POUNAME());

wait();

CASE state OF

  10:

    // arrange: 400 ms period, so the output is high from 200 ms to 400 ms
    pulseTimer.SetPeriod := T#400MS;
    pulseTimer.Signal := TRUE;
    AssertFalse(Condition := pulseTimer.Q_PulseTrain, Message := 'pulse train starts low');
    state := 20;
    wait(IN := TRUE, PT := T#300MS);

  20:

    IF NOT wait.Q THEN
      RETURN;
    END_IF
    wait(IN := FALSE);
    AssertTrue(Condition := pulseTimer.Q_PulseTrain, Message := 'pulse train high in the second half of the period');
    state := 30;
    wait(IN := TRUE, PT := T#200MS);

  30:

    IF NOT wait.Q THEN
      RETURN;
    END_IF
    wait(IN := FALSE);
    AssertFalse(Condition := pulseTimer.Q_PulseTrain, Message := 'pulse train low in the first half of the next period');
    pulseTimer.Signal := FALSE;
    TEST_FINISHED_NAMED(__POUNAME());
    state := 40;

  40:
    ; // finished

END_CASE
END_METHOD

METHOD PRIVATE Test_SetPeriodReadsBackWithMinimumOfOneMs
TcUnit.TEST(__POUNAME());

periodTimer.SetPeriod := T#1S;
AssertEquals_TIME(Expected := T#1S, Actual := periodTimer.SetPeriod, Message := 'period reads back');
periodTimer.SetPeriod := T#0MS;
AssertEquals_TIME(Expected := T#1MS, Actual := periodTimer.SetPeriod, Message := 'period never below 1 ms');

TEST_FINISHED_NAMED(__POUNAME());
END_METHOD

END_FUNCTION_BLOCK

// ---- Tests/T_GetHandle_Tests.TcPOU
// ADS integration: needs the runtime's ADS router (works on the usermode runtime). The suite instance in MAIN must be named suiteGetHandle.
FUNCTION_BLOCK T_GetHandle_Tests EXTENDS TcUnit.FB_TestSuite
VAR
  probe : DINT := 7;
  getHandle : T_GetHandle;
  releaseHandle : T_ReleaseHandle;
  handle : ST_SymbolHandle;
END_VAR

Test_GetsAndReleasesSymbolHandle();

METHOD PRIVATE Test_GetsAndReleasesSymbolHandle
VAR_INST
  state : INT := 10;
  wait : TON;
END_VAR
TcUnit.TEST(__POUNAME());

getHandle();
releaseHandle();
wait();

CASE state OF

  10:

    // arrange: a handle for a symbol of this PLC, over local ADS
    handle.Handle := 0;
    handle.SymbolAddress.SymbolName := 'MAIN.suiteGetHandle.probe';
    handle.SymbolAddress.Ads.port := 851;

    // act
    AssertTrue(Condition := getHandle.TryGetHandle(symbolHandle := handle), Message := 'get handle request accepted');
    state := 20;
    wait(IN := TRUE, PT := T#5S);

  20:

    IF getHandle.Done THEN
      wait(IN := FALSE);
      AssertTrue(Condition := handle.Handle <> 0, Message := 'ADS returned a symbol handle');
      AssertFalse(Condition := getHandle.Busy, Message := 'not busy once done');
      AssertTrue(Condition := releaseHandle.TryReleaseHandle(symbolHandle := handle), Message := 'release handle request accepted');
      state := 30;
      wait(IN := TRUE, PT := T#5S);

    ELSIF getHandle.Error OR wait.Q THEN
      wait(IN := FALSE);
      AssertTrue(Condition := FALSE, Message := 'get handle failed or timed out');
      TEST_FINISHED_NAMED(__POUNAME());
      state := 40;

    END_IF

  30:

    IF releaseHandle.Done THEN
      wait(IN := FALSE);
      AssertFalse(Condition := releaseHandle.Error, Message := 'handle released without error');
      TEST_FINISHED_NAMED(__POUNAME());
      state := 40;

    ELSIF releaseHandle.Error OR wait.Q THEN
      wait(IN := FALSE);
      AssertTrue(Condition := FALSE, Message := 'release handle failed or timed out');
      TEST_FINISHED_NAMED(__POUNAME());
      state := 40;

    END_IF

  40:
    ; // finished

END_CASE
END_METHOD

END_FUNCTION_BLOCK

// ---- Tests/T_InvokeRpcMethod_Tests.TcPOU
// ADS integration: calls an RPC-enabled method of this PLC through ADS. The suite instance in MAIN must be named suiteInvokeRpc.
FUNCTION_BLOCK T_InvokeRpcMethod_Tests EXTENDS TcUnit.FB_TestSuite
VAR
  rpcTarget : T_RpcTarget;
  invoke : T_InvokeRpcMethod;
  addParams : ST_RpcAddParams;
  result : DINT;
  handle : ST_SymbolHandle;
END_VAR

Test_InvokesMethodOverAds();

METHOD PRIVATE Test_InvokesMethodOverAds
VAR_INST
  state : INT := 10;
  wait : TON;
END_VAR
TcUnit.TEST(__POUNAME());

invoke();
wait();

CASE state OF

  10:

    // arrange: call T_RpcTarget.Add on this PLC's own instance through ADS
    addParams.a := 20;
    addParams.b := 22;
    result := 0;
    handle.Handle := 0;
    handle.SymbolAddress.SymbolName := 'MAIN.suiteInvokeRpc.rpcTarget#AddNumbers';
    handle.SymbolAddress.Ads.port := 851;
    handle.SymbolAddress.WriteRef := F_BIGTYPE(pData := ADR(addParams), cbLen := SIZEOF(addParams));
    handle.SymbolAddress.ReadRef := F_BIGTYPE(pData := ADR(result), cbLen := SIZEOF(result));

    // act
    AssertTrue(Condition := invoke.TryInvokeMethodCall(symbolHandle := handle), Message := 'invoke request accepted');
    AssertTrue(Condition := invoke.Busy, Message := 'busy while the call is in flight');
    state := 20;
    wait(IN := TRUE, PT := T#10S);

  20:

    IF invoke.Done THEN
      wait(IN := FALSE);
      AssertEquals_DINT(Expected := 42, Actual := result, Message := 'the RPC method returned a + b');
      AssertEquals_DINT(Expected := 42, Actual := rpcTarget.LastSum, Message := 'the method ran on the target instance');
      AssertFalse(Condition := invoke.Busy, Message := 'not busy once done');
      TEST_FINISHED_NAMED(__POUNAME());
      state := 30;

    ELSIF invoke.Error OR wait.Q THEN
      wait(IN := FALSE);
      AssertTrue(Condition := FALSE, Message := 'ADS RPC call failed or timed out');
      TEST_FINISHED_NAMED(__POUNAME());
      state := 30;

    END_IF

  30:
    ; // finished

END_CASE
END_METHOD

END_FUNCTION_BLOCK

// ---- Mocks/T_RpcTarget.TcPOU
// Target for the ADS RPC tests: AddNumbers is callable through ADS by symbol name.
FUNCTION_BLOCK T_RpcTarget
VAR
  _lastSum : DINT;
END_VAR

{attribute 'TcRpcEnable'}
METHOD AddNumbers : DINT
VAR_INPUT
  a : DINT;
  b : DINT;
END_VAR
AddNumbers := a + b;
_lastSum := AddNumbers;
END_METHOD

PROPERTY LastSum : DINT
GET
LastSum := _lastSum;
END_GET
END_PROPERTY

END_FUNCTION_BLOCK

// ---- Tests/T_WritePersistentData_Tests.TcPOU
FUNCTION_BLOCK T_WritePersistentData_Tests EXTENDS TcUnit.FB_TestSuite

Test_DefaultsToPort851Every10Seconds();
Test_SetConfigChangesPeriodAndPort();
Test_SetConfigRejectsZeroPeriod();
Test_SetConfigRejectsPortZero();

METHOD PRIVATE Test_DefaultsToPort851Every10Seconds
VAR
  persistentWriter : T_WritePersistentData;
END_VAR
TcUnit.TEST(__POUNAME());

AssertEquals_UINT(Expected := 851, Actual := persistentWriter.AdsPort, Message := 'default ADS port');
AssertEquals_TIME(Expected := T#10S, Actual := persistentWriter.WritePeriod, Message := 'default write period');

TEST_FINISHED_NAMED(__POUNAME());
END_METHOD

METHOD PRIVATE Test_SetConfigChangesPeriodAndPort
VAR
  persistentWriter : T_WritePersistentData;
  accepted : BOOL;
END_VAR
TcUnit.TEST(__POUNAME());

accepted := persistentWriter.SetConfig(WritePeriod := T#1M, AdsPort := 852);
AssertTrue(Condition := accepted, Message := 'a period and a port are accepted');
AssertEquals_TIME(Expected := T#1M, Actual := persistentWriter.WritePeriod, Message := 'write period set');
AssertEquals_UINT(Expected := 852, Actual := persistentWriter.AdsPort, Message := 'ADS port set');

TEST_FINISHED_NAMED(__POUNAME());
END_METHOD

METHOD PRIVATE Test_SetConfigRejectsZeroPeriod
VAR
  persistentWriter : T_WritePersistentData;
  accepted : BOOL;
END_VAR
TcUnit.TEST(__POUNAME());

accepted := persistentWriter.SetConfig(WritePeriod := T#0S, AdsPort := 852);
AssertFalse(Condition := accepted, Message := 'a zero period is rejected');
AssertEquals_TIME(Expected := T#10S, Actual := persistentWriter.WritePeriod, Message := 'write period unchanged');
AssertEquals_UINT(Expected := 851, Actual := persistentWriter.AdsPort, Message := 'ADS port unchanged');

TEST_FINISHED_NAMED(__POUNAME());
END_METHOD

METHOD PRIVATE Test_SetConfigRejectsPortZero
VAR
  persistentWriter : T_WritePersistentData;
  accepted : BOOL;
END_VAR
TcUnit.TEST(__POUNAME());

accepted := persistentWriter.SetConfig(WritePeriod := T#1M, AdsPort := 0);
AssertFalse(Condition := accepted, Message := 'port 0 is rejected');
AssertEquals_TIME(Expected := T#10S, Actual := persistentWriter.WritePeriod, Message := 'write period unchanged');
AssertEquals_UINT(Expected := 851, Actual := persistentWriter.AdsPort, Message := 'ADS port unchanged');

TEST_FINISHED_NAMED(__POUNAME());
END_METHOD

END_FUNCTION_BLOCK
